(* IEC 61131-3 sources: Industry-PLC-LLM/data/PLCBEAD_repo/PLCBEAD_PLCEmbed-main/PLC-BEAD/Source/PLC_Programs, 701 files *)

(* ---- NETWORK.IEC ---- *)
(*@PROPERTIES_EX@
TYPE: DATA_TYPE
LOCALE: 0
*)
(*----------------------------------------------------------------------------------*)
TYPE

  oscat_NW_BUF_SHORT : ARRAY [0..1407] OF BYTE;
  oscat_NW_BUF_LONG  : ARRAY [0..4095] OF BYTE;

  oscat_NETWORK_BUFFER_SHORT :
  STRUCT
    SIZE   : UINT;
    BUFFER : oscat_NW_BUF_SHORT;
  END_STRUCT;

  oscat_NETWORK_BUFFER :
  STRUCT
    SIZE   : UINT;
    BUFFER : oscat_NW_BUF_LONG;
  END_STRUCT;

END_TYPE

TYPE oscat_url :
    STRUCT
    PROTOCOL : oscat_STRING10;
    USER     : oscat_STRING32;
    PASSWORD : oscat_STRING32;
    DOMAIN   : oscat_STRING80;
    PORT     : WORD;
    PATH     : oscat_STRING80;
    QUERY    : oscat_STRING250;
    ANCHOR   : oscat_STRING40;
    HEADER   : oscat_STRING160;
    END_STRUCT;
END_TYPE

TYPE
  oscat_aB0_5	: ARRAY [0..5] 	OF BYTE;
  oscat_aB0_15	: ARRAY [0..15]	OF BYTE;
  oscat_aB0_19	: ARRAY [0..19]	OF BYTE;
  oscat_aB0_31	: ARRAY [0..31]	OF BYTE;
  oscat_aB0_39	: ARRAY [0..39]	OF BYTE;
  oscat_aB0_47	: ARRAY [0..47]	OF BYTE;
  oscat_aB0_63	: ARRAY [0..63]	OF BYTE;
  oscat_aB0_255	: ARRAY [0..255] OF BYTE;
  oscat_aB1_255	: ARRAY [1..255] OF BYTE;

  oscat_aW0_255	: ARRAY [0..255] OF WORD;
  oscat_aDW0_3	: ARRAY [0..3] 	OF DWORD;
  oscat_aDW0_15	: ARRAY [0..15] OF DWORD;
  oscat_aDW0_4	: ARRAY [0..4] 	OF DWORD;
  oscat_sDW0_79	: ARRAY [0..79] OF DWORD;
END_TYPE

TYPE
  oscat_VMAP_DATA :
  STRUCT
	FC       : DWORD;
    V_ADR    : INT;
    V_SIZE   : INT;
    P_ADR    : INT;
	TIME_OUT : TIME;
  END_STRUCT;

  oscat_MB_VMAP : ARRAY [1..10] OF oscat_VMAP_DATA;

  csv_parser_demo_col : ARRAY [1..4] OF REAL;
  csv_parser_demo     : ARRAY [1..2] OF csv_parser_demo_col;

END_TYPE

TYPE
  oscat_IP_FIFO128_DATA  : ARRAY [1..128] OF BYTE;
  oscat_Mailbox  : ARRAY [1..16] OF BYTE;

  oscat_IP_FIFO_DATA :
  STRUCT
	X       : oscat_IP_FIFO128_DATA; (* IP_ID FIFO Speicher          *)
	Y       : oscat_IP_FIFO128_DATA; (* IP_ID Z�hler                 *)
	ID      : BYTE;                  (* h�chste vergabene id         *)
	MAX_ID  : BYTE;                  (* maximal Anmeldungen pro ID   *)
    INIT    : BOOL;                  (* Initialisierung durchgef�hrt *)
	EMPTY   : BOOL;                  (* FIFO leer                    *)
	FULL    : BOOL;                  (* FIFO voll                    *)
	TOP     : INT;                   (* maximale anzahl in FIFO      *)
	NW      : INT;                   (* Schreibzeiger                *)
	NR      : INT;                   (* Lesezeiger                   *)
  END_STRUCT;

  oscat_IP_C:
  STRUCT
  	C_MODE:			BYTE;          		(*W Mode: TCP/UCP AKTIV/PASSIV                               *)
	C_PORT:         WORD;          		(*W Portnummer                                               *)
	C_IP:           DWORD;         		(*W IP-Adresse gepackt wwxxyyzz = www.xxx.yyy.zzz            *)
    C_STATE:        BYTE;          		(*R Verbindungsstatus ON/OFF + Flanke ON/OFF                 *)
	C_ENABLE:       BOOL;          		(*W Freigabe f�r Connect                                     *)
    R_OBSERVE:      BOOL;          		(*W Empfang ueberwachen                                      *)
    TIME_RESET:     BOOL;          		(*W Alle Timer ruecksetzen                                   *)
	ERROR:          DWORD;         		(*R vvwwxxyy (vv = CON_ERROR, ww = SEN_ERROR, xx = REC_ERROR *)
    FIFO:           oscat_IP_FIFO_DATA; (*I IP FIFO Struktur                                         *)
	MAILBOX:		oscat_Mailbox;		(*I Mailbox: Datenbereich f�r Bausteindatenaustausch         *)
  END_STRUCT;

  oscat_XML_CONTROL:
  STRUCT
    COMMAND:             WORD;            (*W                 *)
    WATCHDOG:            TIME;            (*W                 *)
    START_POS:           UINT;            (*W                 *)
    STOP_POS:            UINT;            (*W                 *)
    COUNT:               UINT;            (*R                 *)
    TYP:                 INT;             (*R                 *)
    LEVEL:               UINT;            (*R                 *)
    PATH:                oscat_STRING250; (*R                 *)
    ELEMENT:             oscat_STRING250; (*R                 *)
    ATTRIBUTE:           oscat_STRING250; (*R                 *)
    VALUE:               oscat_STRING250; (*R                 *)
    BLOCK1_START:        UINT;            (*R                 *)
    BLOCK1_STOP:         UINT;            (*R                 *)
    BLOCK2_START:        UINT;            (*R                 *)
    BLOCK2_STOP:         UINT;            (*R                 *)
  END_STRUCT;

  (* --------- WORLD WEATHER --------- *)

  oscat_WORLD_WEATHER_CUR :
  STRUCT
	OBSERVATION_TIME : oscat_STRING8;
	TEMP_C           : INT;
	WEATHER_CODE     : INT;
	WEATHER_DESC 	 : oscat_STRING60;
	WEATHER_ICON     : INT;
	WIND_SPEED_MILES : INT;
	WIND_SPEED_KMPH  : INT;
	WIND_DIR_DEGREE  : INT;
	WIND_DIR16POINT  : oscat_STRING3;
	PRECIPMM         : REAL;
	HUMIDITY         : INT;
	VISIBILITY       : INT;
	PRESSURE         : INT;
	CLOUDOVER        : INT;
  END_STRUCT;

  oscat_WORLD_WEATHER_DAY :
  STRUCT
	DATE_OF_DAY      : oscat_STRING10;
	TEMP_MAX_C       : INT;
	TEMP_MAX_F       : INT;
	TEMP_MIN_C       : INT;
	TEMP_MIN_F       : INT;
	WIND_SPEED_MILES : INT;
	WIND_SPEED_KMPH  : INT;
	WIND_DIR_DEGREE  : INT;
	WIND_DIR16POINT  : oscat_STRING3;
	WEATHER_CODE     : INT;
	WEATHER_DESC     : oscat_STRING60;
	WEATHER_ICON     : INT;
	PRECIPMM         : REAL;
  END_STRUCT;

  oscat_WORLD_WEATHER_DAY_ARR : ARRAY [0..4] OF oscat_WORLD_WEATHER_DAY;

  oscat_WORLD_WEATHER_DATA :
  STRUCT
	CUR : oscat_WORLD_WEATHER_CUR;
	DAY : oscat_WORLD_WEATHER_DAY_ARR;
  END_STRUCT;

  oscat_WORLD_WEATHER_aI0_41 : ARRAY[0..41] OF INT;

  (* --------- WEATHER CHANNEL --------- *)
  oscat_YAHOO_WEATHER_DATA:
  STRUCT
    TIMETOLIVE:                 INT;              (* TIME TO LIVE: HOW LONG IN MINUTES THIS FEED SHOULD BE CACHED         *)
    LOCATION_CITY:              OSCAT_STRING40;   (* THE LOCATION OF THIS FORECAST: CITY: CITY NAME  *)
    LOCATION_REGION:            OSCAT_STRING20;   (* THE LOCATION OF THIS FORECAST: REGION: STATE, TERRITORY, OR REGION, IF GIVEN *)
    LOCATION_COUNTRY:           OSCAT_STRING20;    (* THE LOCATION OF THIS FORECAST: COUNTRY: TWO-CHARACTER COUNTRY CODE *)
    UNIT_TEMPERATURE:           OSCAT_STRING1;    (* TEMPERATURE: DEGREE UNITS, F FOR FAHRENHEIT OR C FOR CELSIUS *)
    UNIT_DISTANCE:              OSCAT_STRING2;    (* DISTANCE: UNITS FOR DISTANCE, MI FOR MILES OR KM FOR KILOMETERS *)
    UNIT_PRESSURE:              OSCAT_STRING2;    (* PRESSURE: UNITS OF BAROMETRIC PRESSURE, IN FOR POUNDS PER SQUARE INCH OR MB FOR MILLIBARS *)
    UNIT_SPEED:                 OSCAT_STRING4;    (* SPEED: UNITS OF SPEED, MPH FOR MILES PER HOUR OR KPH FOR KILOMETERS PER HOUR *)
    WIND_CHILL:                 INT;              (* FORECAST INFORMATION ABOUT WIND CHILL IN DEGREES *)
    WIND_DIRECTION:             INT;              (* FORECAST INFORMATION ABOUT WIND DIRECTION, IN DEGREES *)
    WIND_SPEED:                 REAL;             (* FORECAST INFORMATION ABOUT WIND SPEED, IN THE UNITS (MPH OR KPH)*)
    ATMOSPHERE_HUMIDITY:        INT;              (* FORECAST INFORMATION ABOUT CURRENT ATMOSPHERIC HUMIDITY: HUMIDITY, IN PERCENT  *)
    ATMOSPHERE_PRESSURE:        INT;              (* FORECAST INFORMATION ABOUT CURRENT ATMOSPHERIC PRESSURE: BAROMETRIC PRESSURE, IN THE UNITS (IN OR MB) *)
	ATMOSPHERE_VISIBILITY:      REAL;             (* FORECAST INFORMATION ABOUT CURRENT ATMOSPHERIC VISIBILITY, IN THE UNITS (MI OR KM) *)
	ATMOSPHERE_RISING:          INT;              (* FORECAST INFORMATION ABOUT RISING: STATE OF THE BAROMETRIC PRESSURE: STEADY (0), RISING (1), OR FALLING (2). (INTEGER: 0, 1, 2) *)
    ASTRONOMY_SUNRISE:          OSCAT_STRING10;   (* SUNRISE: TODAY'S SUNRISE TIME. THE TIME IS A STRING IN A LOCAL TIME FORMAT OF "H:MM AM/PM" *)
    ASTRONOMY_SUNSET:           OSCAT_STRING10;   (* SUNSET: TODAY'S SUNSET TIME. THE TIME IS A STRING IN A LOCAL TIME FORMAT OF "H:MM AM/PM", *)
    GEO_LATITUDE:               REAL;             (* THE LATITUDE OF THE LOCATION *)
    GEO_LONGITUDE:              REAL;             (* THE LONGITUDE OF THE LOCATION *)
    CUR_CONDITIONS_TEMP:        INT;              (* THE CURRENT WEATHER CONDITIONS: TEMP: THE CURRENT TEMPERATURE, IN THE UNITS (F OR C) *)
    CUR_CONDITIONS_TEXT:        OSCAT_STRING40;   (* THE CURRENT WEATHER CONDITIONS: TEXT: A TEXTUAL DESCRIPTION OF CONDITIONS *)
    CUR_CONDITIONS_CODE:        INT;              (* THE CURRENT WEATHER CONDITIONS: CODE: THE CONDITION CODE FOR THIS FORECAST *)
	CUR_CONDITIONS_ICON:        INT;			  (* THE CURRENT WEATHER CONDITIONS: ICON: THE CONDITION ICON FOR THIS FORECAST *)
    FORCAST_TODAY_LOW_TEMP:     INT;              (* THE FORCAST TODAY WEATHER CONDITIONS: THE FORECASTED LOW TEMPERATURE FOR THIS DAY IN THE UNITS (F OR C) *)
    FORCAST_TODAY_HIGH_TEMP:    INT;              (* THE FORCAST TODAY WEATHER CONDITIONS: THE FORECASTED HIGH TEMPERATURE FOR THIS DAY IN THE UNITS (F OR C) *)
    FORCAST_TODAY_TEXT:         OSCAT_STRING40;   (* THE FORCAST TODAY WEATHER CONDITIONS: TEXT: A TEXTUAL DESCRIPTION OF CONDITIONS *)
    FORCAST_TODAY_CODE:         INT;              (* THE CURRENT WEATHER CONDITIONS: CODE: THE CONDITION CODE FOR THIS FORECAST *)
	FORCAST_TODAY_ICON:         INT;			  (* THE CURRENT WEATHER CONDITIONS: ICON: THE CONDITION ICON FOR THIS FORECAST *)
    FORCAST_TOMORROW_LOW_TEMP:  INT;              (* THE FORCAST TOMORROW WEATHER CONDITIONS: THE FORECASTED LOW TEMPERATURE FOR THIS DAY IN THE UNITS (F OR C) *)
    FORCAST_TOMORROW_HIGH_TEMP: INT;              (* THE FORCAST TOMORROW WEATHER CONDITIONS: THE FORECASTED HIGH TEMPERATURE FOR THIS DAY IN THE UNITS (F OR C) *)
    FORCAST_TOMORROW_TEXT:      OSCAT_STRING40;   (* THE FORCAST TOMORROW WEATHER CONDITIONS: TEXT: A TEXTUAL DESCRIPTION OF CONDITIONS *)
    FORCAST_TOMORROW_CODE:      INT;              (* THE CURRENT WEATHER CONDITIONS: CODE: THE CONDITION CODE FOR THIS FORECAST *)
	FORCAST_TOMORROW_ICON:      INT;			  (* THE CURRENT WEATHER CONDITIONS: ICON: THE CONDITION ICON FOR THIS FORECAST *)
  END_STRUCT;

  oscat_YAHOO_WEATHER_aI0_48 : ARRAY[0..48] OF INT;

  oscat_IP2GEO_DATA:
  STRUCT
	STATE :				BOOL;			  (* STATE *)
	IP4 :				DWORD;			  (* IP-Adresse *)
    COUNTRY_CODE :		oscat_STRING2;    (*   *)
    COUNTRY_NAME :		oscat_STRING20;   (*   *)
    REGION_CODE :		oscat_STRING2;    (*   *)
    REGION_NAME :		oscat_STRING20;   (*   *)
    CITY :				oscat_STRING20;   (*   *)
    GEO_LATITUDE :		REAL;             (*   *)
    GEO_LONGITUDE :		REAL;             (*   *)
	TIME_ZONE_NAME :	oscat_STRING20;
	GMT_OFFSET :		INT;
	IS_DST :			BOOL;
  END_STRUCT;
END_TYPE

(*----------------------------------------------------------------------------------*)

TYPE
  PRINTF_DATA_250  	:  ARRAY [1..11]  OF oscat_STRING250;
  PRINTF_DATA_80 	:  ARRAY [1..11]  OF oscat_STRING80;
  LOG_250       	:  ARRAY [0..400] OF oscat_STRING250;
  LOG_80    		:  ARRAY [0..400] OF oscat_STRING80;
  LOG_OPTION		:  ARRAY [0..400] OF DWORD;

  us_LOG_CONTROL :
  STRUCT
    NEW_MSG              : oscat_STRING250;    (*W neue Nachricht f�r den Datenbuffer   *)
	NEW_MSG_OPTION 		 : DWORD;
    LEVEL                : BYTE;
	SIZE                 : INT;                (*R Anzahl der Strings im LOG_DATA       *)
	RESET                : BOOL;               (*W Nachrichtenbuffer l�schen            *)
    PRINTF               : PRINTF_DATA_250;    (*W Array PRINTF Parameter               *)
    MSG                  : LOG_250;            (*I Array Message                        *)
    MSG_OPTION           : LOG_OPTION;     	   (*I Array Message Option                 *)
	UPDATE_COUNT         : UINT;               (*R Updatez�hler                         *)
    IDX                  : INT;                (*R aktueller Nachrichten-Index          *)
	RING_MODE            : BOOL;               (*I Buffer�berlauf erkannt               *)
  END_STRUCT;

  us_LOG_CONTROL_80 :
  STRUCT
    NEW_MSG              : oscat_STRING80;     (*W neue Nachricht f�r den Datenbuffer   *)
	NEW_MSG_OPTION 		 : DWORD;
    LEVEL                : BYTE;
	SIZE                 : INT;                (*R Anzahl der Strings im LOG_DATA       *)
	RESET                : BOOL;               (*W Nachrichtenbuffer l�schen            *)
    PRINTF               : PRINTF_DATA_80;     (*W Array PRINTF Parameter               *)
    MSG                  : LOG_80;             (*I Array Message                        *)
    MSG_OPTION           : LOG_OPTION;     	   (*I Array Message Option                 *)
	UPDATE_COUNT         : UINT;               (*R Updatez�hler                         *)
    IDX                  : INT;                (*R aktueller Nachrichten-Index          *)
	RING_MODE            : BOOL;               (*I Buffer�berlauf erkannt               *)
  END_STRUCT;

  LINE_ARRAY 			: ARRAY [1..40] OF INT;

  us_LOG_VIEWPORT :
    STRUCT
     LINE_ARRAY          : LINE_ARRAY;
     COUNT               : INT;                (* Anzahl der sichtbaren Nachtrichten   *)
	 UPDATE_COUNT        : UINT;               (* Updatez�hler                         *)
     MOVE_TO_X           : INT;                (* Steuerung der Nachrichtenanzeige     *)
     UPDATE              : BOOL;               (* Daten wurden ge�ndert -> neuzeichnen *)
  END_STRUCT;

  oscat_FILE_SERVER_DATA : STRUCT
	FILE_OPEN	: BOOL;
    FILENAME 	: STRING;
    MODE	 	: BYTE;
    OFFSET   	: UDINT;
    FILE_SIZE   : UDINT;
    AUTO_CLOSE	: TIME;
    ERROR	 	: BYTE;
  END_STRUCT;

  oscat_FILE_PATH_DATA : STRUCT
	DRIVE : oscat_string3;
	DIRECTORY : oscat_string250;
	FILENAME : STRING;
  END_STRUCT;

  oscat_UNI_CIRCULAR_BUFFER_DATA : STRUCT
	D_MODE : INT;
	D_HEAD : WORD;
	D_STRING : oscat_string250;
	D_REAL : REAL;
	D_DWORD : DWORD;
	BUF_SIZE : INT;
	BUF_COUNT : INT;
	BUF_USED : USINT;
	BUF : oscat_NW_BUF_LONG;
	_GetStart : INT;
	_GetEnd : INT;
	_Last : INT;
	_First : INT;
  END_STRUCT;

  oscat_DLOG_DATA : STRUCT
	STORE_TYPE : BYTE;
	ADD_HEADER : BOOL;
	ADD_DATA : BOOL;
	ADD_DATA_REQ : BOOL;
	CLOCK_TRIG : BOOL;
	ID_MAX : USINT;
	DTI : UDINT;
	UCB : oscat_UNI_CIRCULAR_BUFFER_DATA;
	NEW_FILE : STRING;
	NEW_FILE_RTRIG : BOOL;
  END_STRUCT;

END_TYPE
(* --------------------------- NET_VAR ---------------------------- *)
TYPE oscat_NET_VAR_DATA :
STRUCT
	CYCLE : UDINT;
	STATE : BYTE;
	INDEX : INT;
	ID_MAX : USINT;
	ERROR_ID : BYTE;
	BUF_SIZE : UINT;
	S_BUF : oscat_NETWORK_BUFFER;
	R_BUF : oscat_NETWORK_BUFFER;
END_STRUCT;
END_TYPE

TYPE
    oscat_aB1_64 : ARRAY[1..64] OF BYTE;
	oscat_nv_ra : ARRAY[1..8] OF REAL;
	oscat_nv_dw : ARRAY[1..8] OF DWORD;
END_TYPE

(* --------------------------- TELNET ----------------------------- *)

TYPE

(*----------------------------------------------------------------------------------*)
(* Menue-System                                                                     *)
(*----------------------------------------------------------------------------------*)

  us_TN_MENU_POPUP :
  STRUCT
    st_Menu_Text:         oscat_STRING250;   (* X Menue Texte                               *)
    in_Menu_E_Count:      INT;               (*   Menue Elemente Anzahl                     *)
    in_X:                 INT;               (* X Menue X-Position                          *)
    in_Y:                 INT;               (* X Menue Y-Position                          *)
    in_Cols:              INT;               (*   Menue Spaltenanzahl                       *)
    in_Rows:              INT;               (*   Menue Zeilenanzahl                        *)
    in_Cur_Item:          INT;               (* X aktuelles Sub-Menue                       *)
    by_Attr_mF:           BYTE;              (* X Text Attribute mit Fokus                  *)
    by_Attr_oF:           BYTE;              (* X Text Attribute ohne Fokus                 *)
    by_Input_Exten_Code:  BYTE;              (* X Tastencode: Sondertasten                  *)
    bo_Create:            BOOL;              (* X Popup-Menu erzeugen                       *)
    bo_Destroy:           BOOL;              (* X Popup-Menu entfernen                      *)
    bo_Update:            BOOL;              (* X Popup-Menu updaten                        *)
    bo_Activ:             BOOL;              (*   Popup-Menu ist aktiv                      *)
  END_STRUCT;

  us_TN_MENU :
  STRUCT
    st_Menu_Text:         oscat_STRING250;   (* X Menue Texte                               *)
    in_Menu_E_Count:      INT;               (* Menue Elemente Anzahl                       *)
    in_Y:                 INT;               (* Menue Zeilennummer  Y-Position              *)
    in_X:                 INT;               (* Menue Spaltennummer X-Position              *)
    by_Attr_mF:           BYTE;              (* Text Attribute mit Fokus                    *)
    by_Attr_oF:           BYTE;              (* Text Attribute ohne Fokus                   *)
    in_X_SM_new:          INT;               (* neue Sub-Menu X-Position                    *)
    in_Y_SM_new:          INT;               (* neue Sub-Menu Y-Position                    *)
    in_X_SM_old:          INT;               (* alte Sub-Menu X-Position                    *)
    in_Y_SM_old:          INT;               (* alte Sub-Menu Y-Position                    *)
    in_Cur_Menu_Item:     INT;               (* aktuelles Haupt-Menue                       *)
    in_Cur_Sub_Item:      INT;               (* aktuelles Sub-Menue                         *)
    in_State:             INT;               (*   Menu status                               *)
    in_Menu_Selected:     INT;               (* X Menu-Item mit Enter angew�hlt             *)
    bo_Create:            BOOL;              (* X Menu erzeugen                             *)
    bo_Destroy:           BOOL;              (* X Menu entfernen                            *)
    bo_Update:            BOOL;              (* X Menu updaten                              *)

  END_STRUCT;

(*----------------------------------------------------------------------------------*)

  bya_TN_CHAR:       	ARRAY [0..1919] OF BYTE;
  bya_TN_BACKUP:     	ARRAY [0..1919] OF BYTE;
  bya_TN_COLOR:      	ARRAY [0..1919] OF BYTE;
  bya_TN_Line_Update:	ARRAY [0..23]   OF BOOL;

  us_TN_SCREEN :
  STRUCT
    bya_CHAR:			bya_TN_CHAR;
    bya_COLOR:			bya_TN_COLOR;
    bya_BACKUP:			bya_TN_BACKUP;
    bya_Line_Update:	bya_TN_Line_Update;

    by_Input_Exten_Code:    BYTE;
    by_Input_ASCII_Code:    BYTE;
    bo_Input_ASCII_IsNum:   BOOL;
    in_Page_Number:        	INT;                (* aktive Seiten-Nr.              *)
    in_Cursor_X:           	INT;                (* Cursor X-Position              *)
    in_Cursor_Y:           	INT;                (* Cursor Y-Position              *)
    in_EOS_Offset:         	INT;                (* End of String Offset           *)
    by_Clear_Screen_Attr:  	BYTE;               (* Clear-Screen Attr              *)
    bo_Clear_Screen:       	BOOL;               (* Clear-Screen ausl�sen          *)
    bo_Modal_Dialog:       	BOOL;               (* Modaler Dialog ist aktiv       *)
    bo_Menue_Bar_Dialog:   	BOOL;               (* Menue Dialog ist aktiv         *)

  END_STRUCT;

(*----------------------------------------------------------------------------------*)

  us_TN_INPUT_CONTROL_DATA :
  STRUCT
    by_Input_Exten_Code:    BYTE;
    by_Input_ASCII_Code:    BYTE;
    bo_Input_ASCII_IsNum:   BOOL;
    in_Title_X_Offset:  	INT;         	(* Title Text X-Offset                       *)
    in_Title_Y_Offset:   	INT;         	(* Title Text Y-Offset                       *)
    by_Title_Attr:			BYTE;        	(* Title Text Attribute                      *)
    st_Title_String:    	STRING;      	(* Title Text String                         *)
    in_Cursor_X:          	INT;			(* aktuelle Cursor X-Position                *)
    in_Cursor_Y:          	INT;			(* aktuelle Cursor Y-Position                *)
    in_Type:              	INT;            (* Type des Elements                         *)
    in_X:                 	INT;            (* Element X-Position                        *)
    in_Y:                 	INT;            (* Element Y-Position                        *)
    in_Cursor_Pos:        	INT;            (* aktuelle Cursorposition                   *)
    by_Attr_mF:           	BYTE;           (* Text Attribute mit Fokus                  *)
    by_Attr_oF:           	BYTE;           (* Text Attribute ohne Fokus                 *)
	in_selected:          	INT;            (* Text Item wurde ausgew�hlt                *)
    st_Input_Mask:        	STRING;         (* Text Eingabemaske                         *)
    st_Input_Data:        	oscat_STRING250;(* Text aktuelle Eingabedaten                *)
    st_Input_String:      	STRING;         (* Text Kopie nach Return-Taste              *)
    st_Input_ToolTip:     	STRING;         (* Text ToolTip (Eingabeinformation)         *)
	in_Input_Option:      	INT;            (* Text Ausgabe-Optionen                     *)
	bo_Input_Entered:     	BOOL;           (* RETURN-Taste wurde bet�tigt               *)
    bo_Input_Hidden:      	BOOL;           (* Text versteckete Eingabe mit '*'          *)
	bo_Input_Only_Num:    	BOOL;           (* Text nur Nummerneingabe zulassen          *)
	bo_Focus:             	BOOL;           (* Element besitzt den Fokus                 *)
	bo_Update_Input:      	BOOL;           (* Element wegen Benutzereingabe neuzeichnen *)
	bo_Update_All:        	BOOL;           (* Element komplett neuzeichnen              *)

  END_STRUCT;

  usa_TN_INPUT_CONTROL_DATA:   ARRAY [1..20] OF us_TN_INPUT_CONTROL_DATA;

  us_TN_INPUT_CONTROL :
  STRUCT
    bo_Enable:          BOOL;           (* Bearbeitung freigeben/sperren           *)
    bo_Update_all:      BOOL;           (* All Elemente neu zeichnen               *)
    bo_Reset_Fokus:     BOOL;           (* Fokus auf 1. Element setzen             *)
    in_Focus_at:        INT;            (* Controlelement mit aktivem Fokus        *)
    in_Count:           INT;            (* Anzahl der benutzen Control-Elemente    *)
    in_ToolTip_X:       INT;            (* Tooltip Text X-Offset                   *)
    in_ToolTip_Y:		INT;            (* Tooltip Text Y-Offset                   *)
    by_ToolTip_Attr:	BYTE;           (* Tooltip Text Attribute                  *)
    in_ToolTip_Size:	INT;            (* Tooltip Text l�nge                      *)
    usa_TN_INPUT_CONTROL_DATA: usa_TN_INPUT_CONTROL_DATA;
  END_STRUCT;

END_TYPE

(* ---- OSCAT.IEC ---- *)
(*@PROPERTIES_EX@
TYPE: DATA_TYPE
LOCALE: 0
*)
TYPE
  oscat_STRING1               : STRING(1);
  oscat_STRING2               : STRING(2);
  oscat_STRING3               : STRING(3);
  oscat_STRING4               : STRING(4);
  oscat_STRING5               : STRING(5);
  oscat_STRING8               : STRING(8);
  oscat_STRING10              : STRING(10);
  oscat_STRING12              : STRING(12);
  oscat_STRING15              : STRING(15);
  oscat_STRING20              : STRING(20);
  oscat_STRING27              : STRING(27);
  oscat_STRING30              : STRING(30);
  oscat_STRING32              : STRING(32);
  oscat_STRING40              : STRING(40);
  oscat_STRING48              : STRING(48);
  oscat_STRING50              : STRING(50);
  oscat_STRING60              : STRING(60);
  oscat_STRING64              : STRING(64);
  oscat_STRING80              : STRING(80);
  oscat_STRING120             : STRING(120);
  oscat_STRING144             : STRING(144);
  oscat_STRING160             : STRING(160);
  oscat_STRING189             : STRING(189);
  oscat_STRING192             : STRING(192);
  oscat_STRING250             : STRING(250);
END_TYPE

(*----------------------------------------------------------------------------------*)
TYPE

  oscat_arr_0_7               : ARRAY [0..7]    OF REAL;
  oscat_arr_0_15              : ARRAY [0..15]   OF REAL;
  oscat_delay_buf             : ARRAY [0..31]   OF REAL;
  oscat_FT_TN64_array         : ARRAY [0..63]   OF REAL;
  oscat_pt_ARRAY              : ARRAY [1..100]  OF REAL;

  oscat_ardw_0_15             : ARRAY [0..15]   OF DWORD;
  oscat_ardw_0_31             : ARRAY [0..31]   OF DWORD;

  oscat_FILTER_MAV_W          : ARRAY [0..31]   OF WORD;
  oscat_arb_0_3               : ARRAY [0..3]    OF BYTE;

  oscat_esr_collect_data      : ARRAY [0..7]    OF BYTE;
  oscat_DRIVER_4C 			  : ARRAY [1..7] 	OF BYTE;
  oscat_arb_0_249 			  : ARRAY [0..249] 	OF BYTE;
  oscat_bya_LIST_CLEAN        : ARRAY [1..250]  OF BYTE;

  oscat_ari_0_30         	  : ARRAY [0..30]   OF INT;

  oscat_stack_array 		  : ARRAY [1..32]   OF INT;

  oscat_dcf77_bits            : ARRAY [0..58]   OF BOOL;

  oscat_array64_time          : ARRAY [0..63]   OF TIME;

  (* -------------------------------------------------- *)
  oscat_PERIOD2_Y             : ARRAY [0..1]    OF UDINT;
  oscat_PERIOD2_X             : ARRAY [0..3]    OF oscat_PERIOD2_Y;

  oscat_ARRAY_X               : ARRAY [0..1]    OF REAL;
  oscat_XY                    : ARRAY [1..20]   OF oscat_ARRAY_X;

  oscat_parset_X              : ARRAY [1..4]    OF REAL;
  oscat_parset                : ARRAY [0..3]    OF oscat_parset_X;

  oscat_Polynom_ARRAY_X       : ARRAY [0..1]    OF REAL;
  oscat_Polynom_XY            : ARRAY [1..5]    OF oscat_Polynom_ARRAY_X;

END_TYPE

(*----------------------------------------------------------------------------------*)
TYPE oscat_FRACTION :
STRUCT
	NUMERATOR : INT;
	DENOMINATOR : INT;
END_STRUCT;
END_TYPE
(*----------------------------------------------------------------------------------*)
TYPE oscat_CALENDAR :
	STRUCT
		UTC : UDINT;				(* world time UTC *)
		LDT : UDINT;				(* local time *)
		LDATE : UDINT;				(* local date *)
		LTOD : UDINT;				(* local time of day *)
		YEAR : INT;					(* year of LDATE *)
		MONTH : INT;				(* month of LDATE *)
		DAY : INT;					(* day of LDATE *)
		WEEKDAY : INT;				(* weekday of LDATE *)
		OFFSET : INT;				(* Time Zone Offset for Local time in minutes *)
		DST_EN : BOOL;				(* daylight savings time enable *)
		DST_ON : BOOL;				(* true when daylight savings time os on *)
		NAME : oscat_string5;		(* name of time zone *)
		LANGUAGE : INT;			    (* language number pls see language setup *)
		LONGITUDE : REAL;			(* longitude of current location *)
		LATITUDE : REAL;			(* latitude of current location *)
		SUN_RISE : UDINT;			(* sun_rise for current location *)
		SUN_SET : UDINT;			(* sun_set for current location *)
		SUN_MIDDAY : UDINT;			(* worldtime when sun stands at south position *)
		SUN_HEIGTH : REAL;			(* suns heigth at midday, south position *)
		SUN_HOR : REAL;				(* sun angle horizontal 0 = north in degrees *)
		SUN_VER : REAL;				(* sun angle vertical above horizon in degrees *)
		NIGHT : BOOL;				(* true between sun_set and sun_rise *)
		HOLIDAY : BOOL;				(* true when holiday *)
		HOLY_NAME : oscat_string30;	(* name of holiday *)
		WORK_WEEK : INT;			(* current work week *)
	END_STRUCT;
END_TYPE

TYPE oscat_SDT :
STRUCT
	YEAR : INT;
	MONTH : INT;
	DAY : INT;
	WEEKDAY : INT;
	HOUR : INT;
	MINUTE : INT;
	SECOND : INT;
	MS : INT;
END_STRUCT;
END_TYPE

(*----------------------------------------------------------------------------------*)

TYPE oscat_LANGUAGE:
  STRUCT
    DEFAULT 	: INT;
	LMAX    	: INT;
  END_STRUCT;
END_TYPE

(*----------------------------------------------------------------------------------*)
TYPE
	oscat_LOCATION_ELEMENTS	: ARRAY [1..5] OF INT;
END_TYPE

TYPE oscat_LOCATION:
  STRUCT
    DEFAULT 	: INT;
	LMAX    	: INT;
	LANGUAGE	: oscat_LOCATION_ELEMENTS;
  END_STRUCT;
END_TYPE

(*----------------------------------------------------------------------------------*)

TYPE
  oscat_ELEMENT_DIRS 		: ARRAY [0..15] OF oscat_STRING3;
  oscat_DIRS				: ARRAY [1..3]  OF oscat_ELEMENT_DIRS;
END_TYPE

(*----------------------------------------------------------------------------------*)
TYPE
  oscat_CHARNAMES	: ARRAY [1..11] OF STRING;
END_TYPE

(*----------------------------------------------------------------------------------*)

TYPE
  oscat_ELEMENT_MONTHS 	: ARRAY [1..12] OF oscat_STRING10;
  oscat_MONTHS			: ARRAY [1..3]  OF oscat_ELEMENT_MONTHS;
END_TYPE

(*----------------------------------------------------------------------------------*)

TYPE
  oscat_ELEMENT_MONTHS3	: ARRAY [1..12] OF oscat_STRING3;
  oscat_MONTHS3			: ARRAY [1..3]  OF oscat_ELEMENT_MONTHS3;
END_TYPE

(*----------------------------------------------------------------------------------*)

TYPE
  oscat_ELEMENT_WEEKDAYS	: ARRAY [1..7] OF oscat_STRING10;
  oscat_WEEKDAYS			: ARRAY [1..3]  OF oscat_ELEMENT_WEEKDAYS;
END_TYPE

(*----------------------------------------------------------------------------------*)

TYPE
  oscat_ELEMENT_WEEKDAYS2	: ARRAY [1..7] OF oscat_STRING2;
  oscat_WEEKDAYS2			: ARRAY [1..3]  OF oscat_ELEMENT_WEEKDAYS2;
END_TYPE

TYPE oscat_esr_data :
  STRUCT
	typ    : BYTE;
	adress : oscat_string10;
	DS     : UDINT;
	TS     : TIME;
	data   : oscat_esr_collect_data;
  END_STRUCT;
END_TYPE

TYPE
  oscat_ESR_3                : ARRAY [0..3] OF oscat_esr_data;
  oscat_ESR_31               : ARRAY [0..31] OF oscat_esr_data;
END_TYPE

TYPE oscat_vector_3 :
  STRUCT
	X : REAL;
	Y : REAL;
	Z : REAL;
  END_STRUCT;
END_TYPE

TYPE oscat_complex :
  STRUCT
	re : REAL;
	im : REAL;
  END_STRUCT;
END_TYPE

TYPE REAL2 :
  STRUCT
	R1 : REAL;
	RX : REAL;
  END_STRUCT;
END_TYPE

(*----------------------------------------------------------------------------------*)

TYPE oscat_HOLIDAY_DATA :
  STRUCT
	NAME : oscat_string30;
	DAY : SINT;
	MONTH : SINT;
	USE : SINT;
	PAD_BYTE : BYTE;
  END_STRUCT;
END_TYPE

TYPE
  oscat_HOLIDAY_DATA_0_29 	: ARRAY [0..29] OF oscat_HOLIDAY_DATA;
  oscat_HOLIDAY_DATA_0_49 	: ARRAY [0..49] OF oscat_HOLIDAY_DATA;
END_TYPE

(* revision history
hm	18. oct. 2008
	original version

*)

(*	if month = 0 then F_day is the offset in days from easter
	used :0 = NOT used, 1 = used, -1..-7 menas the weekday before the specified DATE example -3 means wednesday before 23.11
*)

(* samples for Holiday data

	HOLIDAY_DE : ARRAY[0..29] OF HOLIDAY_DATA := (name := 'Neujahr', day := 1, month := 1, use := 1),
		(name := 'Heilig Drei Könige', day := 6, month := 1, use := 1),
		(name := 'Karfreitag', day := -2, month := 0, use := 1),
		(name := 'Ostersonntag', day := 0, month := 0, use := 1),
		(name := 'Ostermontag', day := 1, month := 0, use := 1),
		(name := 'Tag der Arbeit', day := 1, month := 5, use := 1),
		(name := 'Christi Himmelfahrt', day := 39, month := 0, use := 1),
		(name := 'Pfingstsonntag', day := 49, month := 0, use := 1),
		(name := 'Pfingstmontag', day := 50, month := 0, use := 1),
		(name := 'Fronleichnam', day := 60, month := 0, use := 1),
		(name := 'Augsburger Friedensfest', day := 8, month := 8, use := 0),
		(name := 'Maria Himmelfahrt', day := 15, month := 8, use := 1),
		(name := 'Tag der Deutschen Einheit', day := 3, month := 10, use := 1),
		(name := 'Reformationstag', day := 31, month := 10, use := 0),
		(name := 'Allerheiligen', day := 1, month := 11, use := 1),
		(name := 'Buss und Bettag', day := 23, month := 11, use := 0),
		(name := '1. Weihnachtstag', day := 25, month := 12, use := 1),
		(name := '2. Weihnachtstag', day := 26, month := 12, use := 1);

	HOLIDAY_AT : ARRAY[0..29] OF HOLIDAY_DATA := (name := 'Neujahr', day := 1, month := 1, use := 1),
		(name := 'Heilig Drei Könige', day := 6, month := 1, use := 1),
		(name := 'Karfreitag', day := -2, month := 0, use := 1),
		(name := 'Ostersonntag', day := 0, month := 0, use := 1),
		(name := 'Ostermontag', day := 1, month := 0, use := 1),
		(name := '', day := 1, month := 5, use := 0),
		(name := 'Christi Himmelfahrt', day := 39, month := 0, use := 1),
		(name := 'Pfingstsonntag', day := 49, month := 0, use := 1),
		(name := 'Pfingstmontag', day := 50, month := 0, use := 1),
		(name := 'Fronleichnam', day := 60, month := 0, use := 1),
		(name := '', day := 8, month := 8, use := 0),
		(name := 'Maria Himmelfahrt', day := 15, month := 8, use := 1),
		(name := '', day := 3, month := 10, use := 0),
		(name := '', day := 31, month := 10, use := 0),
		(name := 'Allerheiligen', day := 1, month := 11, use := 1),
		(name := 'Maria Empfängnis', day := 8, month := 12, use := 1),
		(name := '1. Weihnachtstag', day := 25, month := 12, use := 1),
		(name := '2. Weihnachtstag', day := 26, month := 12, use := 1);

	HOLIDAY_FR : ARRAY[0..29] OF HOLIDAY_DATA := (name := 'Nouvel an', day := 1, month := 1, use := 1),
		(name := 'St Valentin', day := 14, month := 2, use := 0),
		(name := 'Vendredi Saint (alsace)', day := -2, month := 0, use := 0),
		(name := 'Dimanche de pâques', day := 0, month := 0, use := 1),
		(name := 'Lundi de pâques', day := 1, month := 0, use := 1),
		(name := 'Jeudi de Ascension', day := 39, month := 0, use := 1),
		(name := 'dimanche de Pentecôte ', day := 49, month := 0, use := 1),
		(name := 'jeudi de la Trinité', day := 60, month := 0, use := 0),
		(name := 'Fête du travail', day := 1, month := 5, use := 1),
		(name := 'Victoire 1945 ', day := 8, month := 5, use := 1),
		(name := 'Prise de La bastille', day := 14, month := 7, use := 1),
		(name := '15 Août 1944', day := 15, month := 8, use := 1),
		(name := 'Halloween', day := 31, month := 10, use := 0),
		(name := 'Armistice 1918', day := 11, month := 11, use := 1),
		(name := 'Noël', day := 25, month := 12, use := 1),
		(name := 'Saint Étienne (alsace)', day := 26, month := 12, use := 0),
		(name := 'Fête de la musique', day := 21, month := 6, use := 0);

	HOLIDAY_BED : ARRAY[0..29] OF HOLIDAY_DATA :=	(name := 'Neujahr', day := 1, month := 1, use := 1),
		(name := 'Ostersonntag', day := 0, month := 0, use := 1),
		(name := 'Ostermontag', day := 1, month := 0, use := 1),
		(name := 'Tag der Arbeit', day := 1, month := 5, use := 1),
		(name := 'Christi Himmelfahrt', day := 39, month := 0, use := 1),
		(name := 'Pfingsten', day := 49, month := 0, use := 1),
		(name := 'Pfingstmontag', day := 50, month := 0, use := 1),
		(name := 'Nationalfeiertag', day := 21, month := 7, use := 1),
		(name := 'Mariä Himmelfahrt', day := 15, month := 8, use := 1),
		(name := 'Allerheiligen', day := 1, month := 11, use := 1),
		(name := 'Feiertag DG', day := 15, month := 11, use := 1),
		(name := 'Heiligabend', day := 24, month := 12, use := 1),
		(name := '1. Weihnachtstag', day := 25, month := 12, use := 1),
		(name := '2. Weihnachtstag', day := 26, month := 12, use := 1),
		(name := 'Silvester', day := 31, month := 12, use := 1);

	HOLIDAY_ITD : ARRAY[0..29] OF HOLIDAY_DATA := (name := 'Neujahr', day := 1, month := 1, use := 1),
		(name := 'Heilig Drei Könige', day := 6, month := 1, use := 1),
		(name := 'Ostersonntag', day := 0, month := 0, use := 1),
		(name := 'Ostermontag', day := 1, month := 0, use := 1),
		(name := 'Tag der Befeiung Italiens', day := 25, month := 4, use := 1),
		(name := 'Tag der Arbeit', day := 1, month := 5, use := 1),
		(name := 'Pfingsten', day := 49, month := 0, use := 1),
		(name := 'Pfingstmontag', day := 50, month := 0, use := 1),
		(name := 'Tag der Republik Italien', day := 2, month := 6, use := 1),
		(name := 'Mariä Himmelfahrt', day := 15, month := 8, use := 1),
		(name := 'Allerheiligen', day := 1, month := 11, use := 1),
		(name := 'Mariä Empfängnis', day := 8, month := 12, use := 1),
		(name := 'Heiligabend', day := 24, month := 12, use := 0),
		(name := '1. Weihnachtstag', day := 25, month := 12, use := 1),
		(name := '2. Stephanstag', day := 26, month := 12, use := 1);

*)

(* ---- TIMER_P4.ST ---- *)
TYPE oscat_TIMER_EVENT_DATA :
  STRUCT
	TYP          : BYTE;
	CHANNEL      : BYTE;
	DAY          : BYTE;
	START        : UDINT;
	DURATION     : TIME;
	LAND         : BYTE;
	LOR          : BYTE;
	LAST         : UDINT;
  END_STRUCT;
END_TYPE

TYPE
  oscat_TIMER_EVENT           : ARRAY [0..63]    OF oscat_TIMER_EVENT_DATA;
  oscat_TP4_qn                : ARRAY [0..3]    OF BOOL;
END_TYPE

TYPE
  oscat_arb_0_3               : ARRAY [0..3]    OF BYTE;
END_TYPE

FUNCTION _BYTE_TO_INT:INT
	VAR_INPUT
		IN :	BYTE;
	END_VAR

	_BYTE_TO_INT := USINT_TO_INT(BYTE_TO_USINT(IN));
END_FUNCTION

FUNCTION DATE_TO_DT:UDINT
	VAR_INPUT
		IN :	UDINT;
	END_VAR
	DATE_TO_DT := IN;
END_FUNCTION

FUNCTION _DT_TO_DATE_B:UDINT

	VAR_INPUT
		_INN :	UDINT;
	END_VAR

	_DT_TO_DATE_B := (_INN / UDINT#86400) * UDINT#86400;
END_FUNCTION

FUNCTION TIME_TO_UDINT2:UDINT
	VAR_INPUT
		X :	TIME;
	END_VAR

	TIME_TO_UDINT2 := DINT_TO_UDINT(TIME_TO_DINT(X));
END_FUNCTION

FUNCTION DATE_TO_UDINT2:UDINT
	VAR_INPUT
		IN :	UDINT;
	END_VAR

	DATE_TO_UDINT2 := IN;
END_FUNCTION

FUNCTION DAY_OF_WEEK:INT
  VAR_INPUT
    IDATE :	UDINT;
  END_VAR

  DAY_OF_WEEK := UDINT_TO_INT((idate / UDINT#86400 + UDINT#3) MOD UDINT#7) + INT#01;
END_FUNCTION

FUNCTION _BYTE_TO_DINT:DINT
	VAR_INPUT
		IN :	BYTE;
	END_VAR

	_BYTE_TO_DINT := USINT_TO_DINT(BYTE_TO_USINT(IN));
END_FUNCTION

FUNCTION DAY_OF_YEAR_UDINT:INT
	VAR_INPUT
		IDATE :	UDINT;
	END_VAR

	DAY_OF_YEAR_UDINT := UDINT_TO_INT((idate / UDINT#86400) MOD UDINT#1461);
	IF DAY_OF_YEAR_UDINT > 729 THEN
		IF DAY_OF_YEAR_UDINT > 1095 THEN DAY_OF_YEAR_UDINT := DAY_OF_YEAR_UDINT - 1095; ELSE DAY_OF_YEAR_UDINT := DAY_OF_YEAR_UDINT - 729; END_IF;
	ELSIF DAY_OF_YEAR_UDINT > 364 THEN
		DAY_OF_YEAR_UDINT := DAY_OF_YEAR_UDINT - 364;
	ELSE
		DAY_OF_YEAR_UDINT := DAY_OF_YEAR_UDINT + 1;
	END_IF;
END_FUNCTION

FUNCTION MONTH_OF_DATE_UDINT:INT

	VAR_INPUT
		IDATE :	UDINT;
	END_VAR

	MONTH_OF_DATE_UDINT := DAY_OF_YEAR_UDINT(idate);
	IF MONTH_OF_DATE_UDINT < 32 THEN
		MONTH_OF_DATE_UDINT := 1;
	ELSIF LEAP_OF_DATE(IDATE) THEN
		MONTH_OF_DATE_UDINT := (MONTH_OF_DATE_UDINT * 53 + 1668) / 1623;
	ELSE
		MONTH_OF_DATE_UDINT := (MONTH_OF_DATE_UDINT * 53 + 1700) / 1620;
	END_IF;

END_FUNCTION

FUNCTION DAY_OF_MONTH:INT
	VAR_INPUT
		IDATE :	UDINT;
	END_VAR

	day_of_month := day_of_year_UDINT(idate);

	IF leap_of_Date(idate) THEN
		CASE day_of_month OF
			32..60	:	day_of_month := day_of_month - 31;
			61..91	:	day_of_month := day_of_month - 60;
			92..121 :	day_of_month := day_of_month - 91;
			122..152:	day_of_month := day_of_month - 121;
			153..182:	day_of_month := day_of_month - 152;
			183..213:	day_of_month := day_of_month - 182;
			214..244:	day_of_month := day_of_month - 213;
			245..274:	day_of_month := day_of_month - 244;
			275..305:	day_of_month := day_of_month - 274;
			306..335:	day_of_month := day_of_month - 305;
			336..366:	day_of_month := day_of_month - 335;
		END_CASE;
	ELSE
		CASE day_of_month OF
			32..59	:	day_of_month := day_of_month - 31;
			60..90	:	day_of_month := day_of_month - 59;
			91..120 :	day_of_month := day_of_month - 90;
			121..151:	day_of_month := day_of_month - 120;
			152..181:	day_of_month := day_of_month - 151;
			182..212:	day_of_month := day_of_month - 181;
			213..243:	day_of_month := day_of_month - 212;
			244..273:	day_of_month := day_of_month - 243;
			274..304:	day_of_month := day_of_month - 273;
			305..334:	day_of_month := day_of_month - 304;
			335..365:	day_of_month := day_of_month - 334;
		END_CASE;
	END_IF;

END_FUNCTION

FUNCTION LEAP_OF_DATE:BOOL

	VAR_INPUT
		IDATE :	UDINT;
	END_VAR

	LEAP_OF_DATE := SHL(UDINT_TO_DWORD((idate + UDINT#43200) / UDINT#31557600), 30) = DWORD#16#80000000;
END_FUNCTION

FUNCTION DAY_OF_YEAR:INT
	VAR_INPUT
		IDATE :	UDINT;
	END_VAR

	DAY_OF_YEAR := UDINT_TO_INT(((idate) / UDINT#86400) MOD UDINT#1461);
	IF DAY_OF_YEAR > 729 THEN
		IF DAY_OF_YEAR > 1095 THEN DAY_OF_YEAR := DAY_OF_YEAR - 1095; ELSE DAY_OF_YEAR := DAY_OF_YEAR - 729; END_IF;
	ELSIF DAY_OF_YEAR > 364 THEN
		DAY_OF_YEAR := DAY_OF_YEAR - 364;
	ELSE
		DAY_OF_YEAR := DAY_OF_YEAR + 1;
	END_IF;
END_FUNCTION

FUNCTION MONTH_OF_DATE:INT

	VAR_INPUT
		IDATE :	UDINT;
	END_VAR

	MONTH_OF_DATE := DAY_OF_YEAR(idate);
	IF MONTH_OF_DATE < 32 THEN
		MONTH_OF_DATE := 1;
	ELSIF LEAP_OF_DATE((IDATE)) THEN
		MONTH_OF_DATE := (MONTH_OF_DATE * 53 + 1668) / 1623;
	ELSE
		MONTH_OF_DATE := (MONTH_OF_DATE * 53 + 1700) / 1620;
	END_IF;
END_FUNCTION

FUNCTION YEAR_OF_DATE:INT
	VAR_INPUT
		IDATE :	UDINT;
	END_VAR

	YEAR_OF_DATE := UDINT_TO_INT((idate+UDINT#43200) / UDINT#31557600 + UDINT#1970);
END_FUNCTION

FUNCTION _INT_TO_UDINT:UDINT
	VAR_INPUT
		IN :	INT;
	END_VAR

	_INT_TO_UDINT := DINT_TO_UDINT(INT_TO_DINT(IN));
END_FUNCTION

FUNCTION DT_TO_DATE:UDINT
	VAR_INPUT
		IN :	UDINT;
	END_VAR

	DT_TO_DATE := (IN / UDINT#86400) * UDINT#86400;
END_FUNCTION

FUNCTION SET_DT:UDINT

	VAR_INPUT
		YEAR : INT;
		MONTH :	INT;
		DAY : INT;
		HOUR : INT;
		MINUTE : INT;
		SECOND : INT;
	END_VAR

	SET_DT := SET_DATE(YEAR, MONTH, DAY) + _INT_TO_UDINT(SECOND) + _INT_TO_UDINT(MINUTE) * UDINT#60 + _INT_TO_UDINT(HOUR) * UDINT#3600;

END_FUNCTION

FUNCTION SET_DATE:UDINT

	VAR_INPUT
		YEAR :	INT;
		MONTH :	INT;
		DAY :	INT;
	END_VAR

	VAR
		count :	INT;
	END_VAR

	IF month > 2 THEN
		count := (month - 1) * 30;
		IF month > 7 THEN
			count := count + DWORD_TO_INT(SHR(DINT_TO_DWORD(INT_TO_DINT(month) - INT_TO_DINT(3)),1));
		ELSE
			count := count + DWORD_TO_INT(SHR(DINT_TO_DWORD(INT_TO_DINT(month) - INT_TO_DINT(4)),1));
		END_IF;
		IF SHL(INT_TO_WORD(year),14) = WORD#0 THEN
			count := count + 1;
		END_IF;
	ELSE
		count := (month - 1) * 31;
	END_IF;
	SET_DATE := (_INT_TO_UDINT(count + day - 1) + DWORD_TO_UDINT(SHR(UDINT_TO_DWORD(_INT_TO_UDINT(year) * UDINT#1461 - UDINT#2878169), 2))) * UDINT#86400;

END_FUNCTION

FUNCTION MONTH_END:UDINT

	VAR_INPUT
		IDATE :	UDINT;
	END_VAR

	MONTH_END := SET_DATE(YEAR_OF_DATE(idate),MONTH_OF_DATE(idate)+1,1) - UDINT#86400;

END_FUNCTION

FUNCTION YEAR_END:UDINT

	VAR_INPUT
		Y :	INT;
	END_VAR

	YEAR_END := DWORD_TO_UDINT(SHR(UDINT_TO_DWORD(INT_TO_UDINT(y) * UDINT#1461 - UDINT#2876712), 2)) * UDINT#86400;

END_FUNCTION

FUNCTION LEAP_DAY:BOOL

	VAR_INPUT
		IDATE :	UDINT;
	END_VAR

	LEAP_DAY := IDATE MOD UDINT#126230400 = UDINT#68169600;

END_FUNCTION

FUNCTION BIT_LOAD_B:BYTE
	VAR_INPUT
		IN :	BYTE;
		VAL :	BOOL;
		POS :	INT;
	END_VAR

	IF VAL THEN
		BIT_LOAD_B := in OR SHL(BYTE#1,pos);
	ELSE
		BIT_LOAD_B := in AND (NOT SHL(BYTE#1,pos));
	END_IF;
END_FUNCTION

FUNCTION BIT_OF_DWORD : BOOL
  VAR_INPUT
    IN : DWORD;
    N : INT;
  END_VAR

  BIT_OF_DWORD := (SHR(in,N) AND 16#00000001) > 0;
END_FUNCTION

FUNCTION_BLOCK TIMER_P4_Block

	VAR_INPUT
		DTIME :	UDINT;
		TREF_0 :	UDINT;
		TREF_1 :	UDINT;
		HOLY :	BOOL;
		L0 :	BOOL;
		L1 :	BOOL;
		L2 :	BOOL;
		L3 :	BOOL;
		OFS :	BYTE;
		ENQ :	BOOL;
		MAN :	BOOL;
		MI :	BYTE;
		RST :	BOOL;
	END_VAR

	VAR_IN_OUT
		PROG :	oscat_TIMER_EVENT;
	END_VAR

	VAR_OUTPUT
		Q0 :	BOOL;
		Q1 :	BOOL;
		Q2 :	BOOL;
		Q3 :	BOOL;
		STATUS :	BYTE;
	END_VAR

	VAR
		day_start :	UDINT;
		start :	UDINT;
		event :	oscat_TIMER_EVENT_DATA;
		pos :	INT;
		last_execute :	UDINT;
		current_day :	DINT;
		mask :	BYTE;
		ma :	oscat_arb_0_3;
		mo :	oscat_arb_0_3;
		qn :	oscat_TP4_qn;
		qs :	oscat_TP4_qn;
		channel :	INT;
		tx :	UDINT;
		array_max :	INT := 63;
		channel_max :	INT := 3;
	END_VAR

	IF RST THEN
		last_execute := UDINT#00;
		FOR pos := 0 TO ARRAY_MAX DO
			IF (PROG[pos].CHANNEL >= OFS) AND (_BYTE_TO_INT(PROG[pos].CHANNEL) < (_BYTE_TO_INT(OFS) + 4)) THEN PROG[pos].LAST := last_execute; END_IF;
		END_FOR;

		FOR pos := 0 TO channel_max DO
			qs[pos] := FALSE;
		END_FOR;

	ELSIF dtime <> last_execute THEN
		last_execute := DTIME;

		day_start := DATE_TO_DT(_DT_TO_DATE_B(DTIME));

		FOR pos := 0 TO channel_max DO qn[pos] := FALSE; END_FOR;

		FOR pos := 0 TO ARRAY_MAX DO
			event := prog[pos];
			channel := _BYTE_TO_INT(event.CHANNEL) - _BYTE_TO_INT(OFS);
			IF (event.TYP > BYTE#0) AND (channel >= 0) AND (channel <= channel_max) THEN
				ma[channel] := event.LAND;
				mo[channel] := event.LOR;
				CASE _BYTE_TO_INT(event.TYP) OF
					1:
						start := day_start + event.start;
						qn[channel] := dtime >= start AND dtime <= start + TIME_TO_UDINT2(event.DURATION);

					2:
						IF (SHR(BYTE#128, DAY_OF_WEEK(_DT_TO_DATE_B(Dtime))) AND event.DAY) > BYTE#0 THEN
							start := day_start + event.start;
							qn[channel] := dtime >= start AND dtime <= start + TIME_TO_UDINT2(event.DURATION);
						END_IF;

					3:
						IF current_day MOD _BYTE_TO_DINT(event.DAY) = DINT#0 THEN
							start := day_start + event.start;
							qn[channel] := dtime >= start AND dtime <= start + TIME_TO_UDINT2(event.DURATION);
						END_IF;

					10:
						IF DAY_OF_WEEK(_DT_TO_DATE_B(DTIME)) = BYTE_TO_INT(event.DAY) THEN
							start := day_start + event.start;
							qn[channel] := dtime >= start AND dtime <= start + TIME_TO_UDINT2(event.DURATION);
						END_IF;

					20:
						IF DAY_OF_MONTH(_DT_TO_DATE_B(DTIME)) = BYTE_TO_INT(event.DAY) THEN
							start := day_start + event.start;
							qn[channel] := dtime >= start AND dtime <= start + TIME_TO_UDINT2(event.DURATION);
						END_IF;

					21:
						IF _DT_TO_DATE_B(DTIME) = MONTH_END(_DT_TO_DATE_B(dtime)) THEN
							start := day_start + event.start;
							qn[channel] := dtime >= start AND dtime <= start + TIME_TO_UDINT2(event.DURATION);
						END_IF;

					30:
						IF DAY_OF_YEAR(_DT_TO_DATE_B(DTIME)) = BYTE_TO_INT(event.DAY) THEN
							start := day_start + event.start;
							qn[channel] := dtime >= start AND dtime <= start + TIME_TO_UDINT2(event.DURATION);
						END_IF;

					31:
						IF _DT_TO_DATE_B(DTIME) = YEAR_END(YEAR_OF_DATE(_DT_TO_DATE_B(dtime))) THEN
							start := day_start + event.start;
							qn[channel] := dtime >= start AND dtime <= start + TIME_TO_UDINT2(event.DURATION);
						END_IF;

					40:
						IF LEAP_DAY(_DT_TO_DATE_B(dtime)) THEN
							start := day_start + event.start;
							qn[channel] := dtime >= start AND dtime <= start + TIME_TO_UDINT2(event.DURATION);
						END_IF;

					41:
						IF HOLY THEN
							start := day_start + event.start;
							qn[channel] := dtime >= start AND dtime <= start + TIME_TO_UDINT2(event.DURATION);
						END_IF;

					42:
						IF (Holy OR (DAY_OF_WEEK(_DT_TO_DATE_B(dtime)) = 6) OR (DAY_OF_WEEK(_DT_TO_DATE_B(dtime)) = 7)) THEN
							start := day_start + event.start;
							qn[channel] := dtime >= start AND dtime <= start + TIME_TO_UDINT2(event.DURATION);
						END_IF;

					43:
						IF DAY_OF_WEEK(_DT_TO_DATE_B(dtime)) < 6 THEN
							start := day_start + event.start;
							qn[channel] := dtime >= start AND dtime <= start + TIME_TO_UDINT2(event.DURATION);
						END_IF;

					50:
						CASE _BYTE_TO_INT(prog[pos].DAY) OF
							0:	tx := tref_0;
							1:	tx := tref_1;
						ELSE
							tx := UDINT#0 ;
						END_CASE;
						start := day_start + tx + event.start;
						qn[channel] := dtime >= start AND dtime <= start + TIME_TO_UDINT2(event.DURATION);

					51:
						CASE _BYTE_TO_INT(prog[pos].DAY) OF
							0:	tx := tref_0;
							1:	tx := tref_1;
						ELSE
							tx := UDINT#0;
						END_CASE;
						start := day_start + tx - event.start;
						qn[channel] := dtime >= start AND dtime <= start + TIME_TO_UDINT2(event.DURATION);

					52 :
						CASE _BYTE_TO_INT(prog[pos].DAY) OF
							0:	tx := tref_0;
							1:	tx := tref_1;
						ELSE
							tx := UDINT#0 ;
						END_CASE;
						start := day_start + tx + event.start;
						IF dtime >= start AND day_start > event.LAST THEN
							qs[channel] := TRUE;
							prog[pos].LAST := day_start;
						END_IF;

					53 :
						CASE _BYTE_TO_INT(prog[pos].DAY) OF
							0:	tx := tref_0;
							1:	tx := tref_1;
						ELSE
							tx := UDINT#0 ;
						END_CASE;
						start := day_start + tx + event.start;
						IF dtime >= start AND day_start > event.LAST THEN
							qs[channel] := FALSE;
							prog[pos].LAST := day_start;
						END_IF;

					54 :
						CASE _BYTE_TO_INT(prog[pos].DAY) OF
							0:	tx := tref_0;
							1:	tx := tref_1;
						ELSE
							tx := UDINT#0 ;
						END_CASE;
						start := day_start + tx - event.start;
						IF dtime >= start AND day_start > event.LAST THEN
							qs[channel] := TRUE;
							prog[pos].LAST := day_start;
						END_IF;

					55 :
						CASE _BYTE_TO_INT(prog[pos].DAY) OF
							0:	tx := tref_0;
							1:	tx := tref_1;
						ELSE
							tx := UDINT#0 ;
						END_CASE;
						start := day_start + tx - event.start;
						IF dtime >= start AND day_start > event.LAST THEN
							qs[channel] := FALSE;
							prog[pos].LAST := day_start;
						END_IF;
				END_CASE;
			END_IF;
		END_FOR;
	END_IF;

	mask := BYTE#255;
	mask:=BIT_LOAD_B(mask,L0,0);
	mask:=BIT_LOAD_B(mask,L1,1);
	mask:=BIT_LOAD_B(mask,L2,2);
	mask:=BIT_LOAD_B(mask,L3,3);

	Q0 := ENQ AND ((qn[0] OR qs[0]) AND ((ma[0] AND mask) = ma[0]) OR ((mo[0] AND mask) > BYTE#0) OR (man AND BIT_OF_DWORD(BYTE_TO_DWORD(MI),0)));
	Q1 := ENQ AND ((qn[1] OR qs[1]) AND ((ma[1] AND mask) = ma[1]) OR ((mo[1] AND mask) > BYTE#1) OR (man AND BIT_OF_DWORD(BYTE_TO_DWORD(MI),1)));
	Q2 := ENQ AND ((qn[2] OR qs[2]) AND ((ma[2] AND mask) = ma[2]) OR ((mo[2] AND mask) > BYTE#2) OR (man AND BIT_OF_DWORD(BYTE_TO_DWORD(MI),2)));
	Q3 := ENQ AND ((qn[3] OR qs[3]) AND ((ma[3] AND mask) = ma[3]) OR ((mo[3] AND mask) > BYTE#3) OR (man AND BIT_OF_DWORD(BYTE_TO_DWORD(MI),3)));

	IF NOT enq THEN
		status := BYTE#100;
	ELSIF man THEN
		status := BYTE#101;
	ELSE
		status := BYTE#102;
	END_IF;

END_FUNCTION_BLOCK

PROGRAM program0
	VAR
		DTIME :	UDINT;
		TREF_0 :	UDINT;
		TREF_1 :	UDINT;
		HOLY :	BOOL;
		L0 :	BOOL;
		L1 :	BOOL;
		L2 :	BOOL;
		L3 :	BOOL;
		OFS :	BYTE;
		ENQ :	BOOL;
		MAN :	BOOL;
		MI :	BYTE;
		RST :	BOOL;
		PROG :	oscat_TIMER_EVENT;
		Q0 :	BOOL;
		Q1 :	BOOL;
		Q2 :	BOOL;
		Q3 :	BOOL;
		STATUS :	BYTE;

		func_block : TIMER_P4_Block;
	END_VAR
	func_block.DTIME := DTIME;
	func_block.TREF_0 := TREF_0;
	func_block.TREF_1 := TREF_1;
	func_block.HOLY := HOLY;
	func_block.L0 := L0;
	func_block.L1 := L1;
	func_block.L2 := L2;
	func_block.L3 := L3;
	func_block.OFS := OFS;
	func_block.ENQ := ENQ;
	func_block.MAN := MAN;
	func_block.MI := MI;
	func_block.RST := RST;
	func_block.PROG := PROG;

	func_block();
	PROG  := func_block.PROG;
	Q0  := func_block.Q0;
	Q1  := func_block.Q1;
	Q2  := func_block.Q2;
	Q3  := func_block.Q3;
	STATUS  := func_block.STATUS;
END_PROGRAM

CONFIGURATION Config0
	RESOURCE Res0 ON PLC
		TASK task0(INTERVAL := T#20ms,PRIORITY := 0);
		PROGRAM instance0 WITH task0 : program0;
	END_RESOURCE
END_CONFIGURATION

(* ---- WORLD_WEATHER.ST ---- *)
TYPE
  oscat_STRING30              : STRING;
  oscat_STRING250             : STRING;
  oscat_STRING8               : STRING;
  oscat_STRING60               : STRING;
  oscat_STRING3               : STRING;
  oscat_STRING10               : STRING;
END_TYPE

TYPE
  oscat_IP_FIFO128_DATA  : ARRAY [1..128] OF BYTE;
  oscat_Mailbox  : ARRAY [1..16] OF BYTE;

  oscat_IP_FIFO_DATA :
  STRUCT
	X       : oscat_IP_FIFO128_DATA; (* IP_ID FIFO Speicher          *)
	Y       : oscat_IP_FIFO128_DATA; (* IP_ID Z�hler                 *)
	ID      : BYTE;                  (* h�chste vergabene id         *)
	MAX_ID  : BYTE;                  (* maximal Anmeldungen pro ID   *)
    INIT    : BOOL;                  (* Initialisierung durchgef�hrt *)
	EMPTY   : BOOL;                  (* FIFO leer                    *)
	FULL    : BOOL;                  (* FIFO voll                    *)
	TOP     : INT;                   (* maximale anzahl in FIFO      *)
	NW      : INT;                   (* Schreibzeiger                *)
	NR      : INT;                   (* Lesezeiger                   *)
  END_STRUCT;

  oscat_IP_C:
  STRUCT
  	C_MODE:			BYTE;          		(*W Mode: TCP/UCP AKTIV/PASSIV                               *)
	C_PORT:         WORD;          		(*W Portnummer                                               *)
	C_IP:           DWORD;         		(*W IP-Adresse gepackt wwxxyyzz = www.xxx.yyy.zzz            *)
    C_STATE:        BYTE;          		(*R Verbindungsstatus ON/OFF + Flanke ON/OFF                 *)
	C_ENABLE:       BOOL;          		(*W Freigabe f�r Connect                                     *)
    R_OBSERVE:      BOOL;          		(*W Empfang ueberwachen                                      *)
    TIME_RESET:     BOOL;          		(*W Alle Timer ruecksetzen                                   *)
	ERROR:          DWORD;         		(*R vvwwxxyy (vv = CON_ERROR, ww = SEN_ERROR, xx = REC_ERROR *)
    FIFO:           oscat_IP_FIFO_DATA; (*I IP FIFO Struktur                                         *)
	MAILBOX:		oscat_Mailbox;		(*I Mailbox: Datenbereich f�r Bausteindatenaustausch         *)
  END_STRUCT;

  oscat_XML_CONTROL:
  STRUCT
    COMMAND:             WORD;            (*W                 *)
    WATCHDOG:            TIME;            (*W                 *)
    START_POS:           UINT;            (*W                 *)
    STOP_POS:            UINT;            (*W                 *)
    COUNT:               UINT;            (*R                 *)
    TYP:                 INT;             (*R                 *)
    LEVEL:               UINT;            (*R                 *)
    PATH:                oscat_STRING250; (*R                 *)
    ELEMENT:             oscat_STRING250; (*R                 *)
    ATTRIBUTE:           oscat_STRING250; (*R                 *)
    VALUE:               oscat_STRING250; (*R                 *)
    BLOCK1_START:        UINT;            (*R                 *)
    BLOCK1_STOP:         UINT;            (*R                 *)
    BLOCK2_START:        UINT;            (*R                 *)
    BLOCK2_STOP:         UINT;            (*R                 *)
  END_STRUCT;

  (* --------- WORLD WEATHER --------- *)

  oscat_WORLD_WEATHER_CUR :
  STRUCT
	OBSERVATION_TIME : oscat_STRING8;
	TEMP_C           : INT;
	WEATHER_CODE     : INT;
	WEATHER_DESC 	 : oscat_STRING60;
	WEATHER_ICON     : INT;
	WIND_SPEED_MILES : INT;
	WIND_SPEED_KMPH  : INT;
	WIND_DIR_DEGREE  : INT;
	WIND_DIR16POINT  : oscat_STRING3;
	PRECIPMM         : REAL;
	HUMIDITY         : INT;
	VISIBILITY       : INT;
	PRESSURE         : INT;
	CLOUDOVER        : INT;
  END_STRUCT;

  oscat_WORLD_WEATHER_DAY :
  STRUCT
	DATE_OF_DAY      : oscat_STRING10;
	TEMP_MAX_C       : INT;
	TEMP_MAX_F       : INT;
	TEMP_MIN_C       : INT;
	TEMP_MIN_F       : INT;
	WIND_SPEED_MILES : INT;
	WIND_SPEED_KMPH  : INT;
	WIND_DIR_DEGREE  : INT;
	WIND_DIR16POINT  : oscat_STRING3;
	WEATHER_CODE     : INT;
	WEATHER_DESC     : oscat_STRING60;
	WEATHER_ICON     : INT;
	PRECIPMM         : REAL;
  END_STRUCT;

  oscat_WORLD_WEATHER_DAY_ARR : ARRAY [0..4] OF oscat_WORLD_WEATHER_DAY;

  oscat_WORLD_WEATHER_DATA :
  STRUCT
	CUR : oscat_WORLD_WEATHER_CUR;
	DAY : oscat_WORLD_WEATHER_DAY_ARR;
  END_STRUCT;

  oscat_WORLD_WEATHER_aI0_41 : ARRAY[0..41] OF INT;

END_TYPE

TYPE
  oscat_NW_BUF_LONG  : ARRAY [0..4095] OF BYTE;

  oscat_NETWORK_BUFFER :
  STRUCT
    SIZE   : UINT;
    BUFFER : oscat_NW_BUF_LONG;
  END_STRUCT;

END_TYPE

FUNCTION_BLOCK WORLD_WEATHER_Block

	VAR_INPUT
		ACTIVATE :	BOOL;
		LATITUDE :	REAL;
		LONGITUDE :	REAL;
		KEY :	oscat_STRING30;
	END_VAR

	VAR_OUTPUT
		BUSY :	BOOL;
		DONE :	BOOL;
		ERROR_C :	DWORD;
		ERROR_T :	BYTE;
	END_VAR

	VAR_IN_OUT
		IP_C :	oscat_IP_C;
		S_BUF :	oscat_NETWORK_BUFFER;
		R_BUF :	oscat_NETWORK_BUFFER;
		WW :	oscat_WORLD_WEATHER_DATA;
	END_VAR

	VAR
		CHK_REAL :	CHK_REAL;
		REAL_TO_STRF :	REAL_TO_STRF;
		URL_DATA :	oscat_url;
		DNS_CLIENT :	DNS_CLIENT;
		HTTP_GET :	HTTP_GET;
		CPB :	CSV_PARSER_BUF;
		STRING_TO_URL :	STRING_TO_URL;
		FLOAT_TO_REAL :	FLOAT_TO_REAL;
		last_state :	BOOL;
		value_int :	INT;
		value_real :	REAL;
		v_real :	REAL;
		state :	INT;
		url_str :	oscat_STRING250;
		offset :	UDINT;
		size :	INT;
		sep :	BYTE;
		cnt :	INT;
		day :	INT;
		idx :	INT;
		run :	BYTE;
		result :	BYTE;
		value :	oscat_STRING250;
		DEC_TO_INT :	DEC_TO_INT;
		pos :	INT;
	END_VAR

	CASE state OF

	00:
		IF ACTIVATE AND NOT last_state THEN
			state := 20;
			DONE := FALSE;
			BUSY := TRUE;
			ERROR_C := DWORD#0;
			ERROR_T := BYTE#0;
		END_IF;

	20:
		REAL_TO_STRF(IN:=LATITUDE,N:=6,D:='.');
		url_str := CONCAT('http://free.worldweatheronline.com/feed/weather.ashx?q=',REAL_TO_STRF.REAL_TO_STRF);
		url_str := CONCAT(url_str,',');
		REAL_TO_STRF(IN:=LONGITUDE,N:=6,D:='.');
		url_str := CONCAT(url_str,REAL_TO_STRF.REAL_TO_STRF);
		url_str := CONCAT(url_str,'&format=csv&num_of_days=5&key=');
		url_str := CONCAT(url_str,key);

		STRING_TO_URL(STR:=url_str, DEFAULT_PROTOCOL:='', DEFAULT_PATH:='' );
		URL_DATA:=STRING_TO_URL.STRING_TO_URL;

		state := 40;

	40:
		IF DNS_CLIENT.DONE THEN
			state := 60;
		ELSIF (DNS_CLIENT.ERROR > DWORD#00) THEN
			ERROR_C := DNS_CLIENT.ERROR;
			ERROR_T := BYTE#01;
			state   := 100;
		END_IF;

	60:
		IF HTTP_GET.DONE THEN
			sep := BYTE#0;
			idx := 0;
			day := 0;
			cnt := 0;
			OFFSET := UINT_TO_UDINT(HTTP_GET.BODY_START);
			size := UINT_TO_INT(HTTP_GET.BODY_STOP);
			run := BYTE#1;
			state := 80;

		ELSIF (HTTP_GET.ERROR > DWORD#00) THEN
			ERROR_C := HTTP_GET.ERROR;
			ERROR_T := BYTE#02;
			state := 100;
		END_IF;

	80:	IF run = BYTE#0 THEN
			run := BYTE#1;
			IF result = BYTE#1 OR result = BYTE#2 THEN
				value_int := 0;
				value_real := 0.0;
				IF LEN(value) <= 20 THEN
					FLOAT_TO_REAL(FLT:=value);
					v_real := FLOAT_TO_REAL.FLOAT_TO_REAL;
					CHK_REAL(X := v_real);
					IF CHK_REAL.CHK_REAL = BYTE#0 THEN
						value_real := v_real;
						value_int := REAL_TO_INT(value_real);
					END_IF;
				END_IF;
				cnt := cnt + 1;
				IF cnt >=8 AND cnt <= 87 THEN
					IF cnt > 22 THEN
						CASE idx OF
						00:	WW.DAY[day].DATE_OF_DAY := value;
						01:	WW.DAY[day].TEMP_MAX_C := value_int;
						02:	WW.DAY[day].TEMP_MAX_F := value_int;
						03:	WW.DAY[day].TEMP_MIN_C := value_int;
						04:	WW.DAY[day].TEMP_MIN_F := value_int;
						05:	WW.DAY[day].WIND_SPEED_MILES := value_int;
						06:	WW.DAY[day].WIND_SPEED_KMPH := value_int;
						07:	WW.DAY[day].WIND_DIR_DEGREE := value_int;
						08:	WW.DAY[day].WIND_DIR16POINT := value;
						09:	WW.DAY[day].WEATHER_CODE := value_int;
						10:	pos := FIND(value, '/wsymbol_');
							IF pos > 0 AND LEN(value) > pos + 13 THEN
								DEC_TO_INT(DEC:=MID(value,4,pos + 9));
								WW.DAY[day].WEATHER_ICON := DEC_TO_INT.DEC_TO_INT;
							ELSE
								WW.DAY[day].WEATHER_ICON := 0;
							END_IF;
						11:	WW.DAY[day].WEATHER_DESC := value;
						12:	WW.DAY[day].PRECIPMM := value_real;
						END_CASE;
						idx := idx + 1;
						IF idx > 12 THEN
							idx := 0;
							day := day + 1;
						END_IF;
					ELSE
						CASE cnt OF
						08:	sep := BYTE#44;
						09:	WW.CUR.OBSERVATION_TIME := value;
						10:	WW.CUR.TEMP_C := value_int;
						11:	WW.CUR.WEATHER_CODE := value_int;
						12:	pos := FIND(value, '/wsymbol_');
							IF pos > 0 AND LEN(value) > pos + 13 THEN
								DEC_TO_INT(DEC:=MID(value,4,pos + 9));
								WW.CUR.WEATHER_ICON := DEC_TO_INT.DEC_TO_INT;
							ELSE
								WW.CUR.WEATHER_ICON := 0;
							END_IF;
						13:	WW.CUR.WEATHER_DESC := value;
						14:	WW.CUR.WIND_SPEED_MILES := value_int;
						15:	WW.CUR.WIND_SPEED_KMPH := value_int;
						16:	WW.CUR.WIND_DIR_DEGREE := value_int;
						17:	WW.CUR.WIND_DIR16POINT := value;
						18:	WW.CUR.PRECIPMM := value_real;
						19:	WW.CUR.HUMIDITY := value_int;
						20:	WW.CUR.VISIBILITY := value_int;
						21:	WW.CUR.PRESSURE := value_int;
						22:	WW.CUR.CLOUDOVER := value_int;
						END_CASE;
					END_IF;
				END_IF;
			ELSIF result = BYTE#10 THEN
				DONE  := TRUE;
				run := BYTE#0;
				state := 100;
			END_IF;
		END_IF;

	100:
		IF (NOT HTTP_GET.DONE) THEN
			state := 0;
			BUSY := FALSE;
			DONE := ERROR_T = BYTE#0;
		END_IF;

	END_CASE;

	DNS_CLIENT.IP_C     := IP_C;
	DNS_CLIENT.S_BUF    := S_BUF;
	DNS_CLIENT.R_BUF    := R_BUF;
	DNS_CLIENT.DOMAIN   := URL_DATA.DOMAIN;
	DNS_CLIENT.IP4_DNS  := DWORD#00;
	DNS_CLIENT.ACTIVATE := state=40;
	DNS_CLIENT();
	IP_C  := DNS_CLIENT.IP_C;
	S_BUF := DNS_CLIENT.S_BUF;
	R_BUF := DNS_CLIENT.R_BUF;

	HTTP_GET.IP_C        := IP_C;
	HTTP_GET.S_BUF       := S_BUF;
	HTTP_GET.R_BUF       := R_BUF;
	HTTP_GET.IP4         := DNS_CLIENT.IP4;
	HTTP_GET.GET         := state=60;
	HTTP_GET.MODE        := BYTE#2;
	HTTP_GET.UNLOCK_BUF  := state=100;
	HTTP_GET.URL_DATA    := URL_DATA;
	HTTP_GET();
	IP_C     := HTTP_GET.IP_C;
	S_BUF    := HTTP_GET.S_BUF;
	R_BUF    := HTTP_GET.R_BUF;
	URL_DATA := HTTP_GET.URL_DATA;

	CPB(SEP:=sep,RUN:=run,OFFSET:=offset,VALUE:=value,PT:=R_BUF);
	run:=CPB.RUN;
	offset:=CPB.OFFSET;
	value:=CPB.VALUE;
	R_BUF:=CPB.PT;
	result:=CPB.RESULT;

	last_state := ACTIVATE;

END_FUNCTION_BLOCK

PROGRAM program0
	VAR
		ACTIVATE :	BOOL;
		LATITUDE :	REAL;
		LONGITUDE :	REAL;
		KEY :	oscat_STRING30;
		IP_C :	oscat_IP_C;
		S_BUF :	oscat_NETWORK_BUFFER;
		R_BUF :	oscat_NETWORK_BUFFER;
		WW :	oscat_WORLD_WEATHER_DATA;
		BUSY :	BOOL;
		DONE :	BOOL;
		ERROR_C :	DWORD;
		ERROR_T :	BYTE;

		func_block : WORLD_WEATHER_Block;
	END_VAR
	func_block.ACTIVATE := ACTIVATE;
	func_block.LATITUDE := LATITUDE;
	func_block.LONGITUDE := LONGITUDE;
	func_block.KEY := KEY;
	func_block.IP_C := IP_C;
	func_block.S_BUF := S_BUF;
	func_block.R_BUF := R_BUF;
	func_block.WW := WW;

	func_block();
	IP_C  := func_block.IP_C;
	S_BUF  := func_block.S_BUF;
	R_BUF  := func_block.R_BUF;
	WW  := func_block.WW;
	BUSY  := func_block.BUSY;
	DONE  := func_block.DONE;
	ERROR_C  := func_block.ERROR_C;
	ERROR_T  := func_block.ERROR_T;
END_PROGRAM

CONFIGURATION Config0
	RESOURCE Res0 ON PLC
		TASK task0(INTERVAL := T#20ms,PRIORITY := 0);
		PROGRAM instance0 WITH task0 : program0;
	END_RESOURCE
END_CONFIGURATION

(* ---- A_TRIG.ST ---- *)
FUNCTION_BLOCK A_TRIG

	VAR_INPUT
		IN :	REAL;
		RES :	REAL;
	END_VAR

	VAR_OUTPUT
		Q :	BOOL;
		D :	REAL;
	END_VAR

	VAR
		last_in :	REAL;
	END_VAR

	D := IN - LAST_IN;
	IF ABS(D) >= res THEN
		Q := TRUE;
		last_in := IN;
	ELSE
		Q := FALSE;
	END_IF;

END_FUNCTION_BLOCK

PROGRAM program0
	VAR
	    LocalVar0 : REAL;
		LocalVar1 : REAL;
		LocalOUT1  : BOOL;
		LocalOUT2  : REAL;
		func_block : A_TRIG;
  	END_VAR
	func_block.IN := LocalVar0;
    func_block.RES := LocalVar1;
	func_block();
	LocalOUT1 := func_block.Q;
	LocalOUT2 := func_block.D;
END_PROGRAM

CONFIGURATION Config0
  	RESOURCE Res0 ON PLC
    	TASK task0(INTERVAL := T#20ms,PRIORITY := 0);
    	PROGRAM instance0 WITH task0 : program0;
  	END_RESOURCE
END_CONFIGURATION

(* ---- ACTUATOR_2P.ST ---- *)
FUNCTION UDINT_TO_TIME2:TIME

	VAR_INPUT
		IN :	UDINT;
	END_VAR

	UDINT_TO_TIME2 := DINT_TO_TIME(UDINT_TO_DINT(IN));

END_FUNCTION

FUNCTION_BLOCK T_PLC_MS_block
	VAR_OUTPUT
		T_PLC_MS :	UDINT;
	END_VAR

	VAR_EXTERNAL
		PLC_TICKS_PER_SEC :	INT;
		PLC_SYS_TICK_CNT :	DINT;
	END_VAR

	VAR
		debug :	BOOL;(*Debug-Mode ON / OFF*)
		N :	INT;(*Debug-Faktor*)
		Offset :	UDINT;(*Debug-Offset*)
		temp :	DWORD := DWORD#1;(*Debug-Offset*)
		mode :	BOOL;(*modus*)
		faktor :	UDINT;(*Systemtakt-Faktor*)
		init :	BOOL;
		v_plc_ticks_per_sec :	UDINT;
		base :	UDINT := UDINT#1000;
	END_VAR

	IF init = FALSE THEN
		v_plc_ticks_per_sec := INT_TO_UDINT(PLC_TICKS_PER_SEC);
		IF v_plc_ticks_per_sec = UDINT#1024 THEN
			faktor := UDINT#1;
			mode := FALSE;
		ELSIF v_plc_ticks_per_sec > UDINT#0 THEN
			IF v_plc_ticks_per_sec <= base THEN
				faktor := base / v_plc_ticks_per_sec;
				mode := FALSE;
			ELSE
				faktor := v_plc_ticks_per_sec / base;
				mode := TRUE;
			END_IF;
		ELSE
			faktor := UDINT#1;
		END_IF;
		init := TRUE;
	END_IF;

	IF mode THEN
		T_PLC_MS := DINT_TO_UDINT(PLC_SYS_TICK_CNT) / faktor;
	ELSE
		T_PLC_MS := DINT_TO_UDINT(PLC_SYS_TICK_CNT) * faktor;
	END_IF;

	IF debug THEN
		T_PLC_MS := (DWORD_TO_UDINT(SHL(UDINT_TO_DWORD(T_PLC_MS),N) OR SHL(temp,N)) - UDINT#1) + Offset;
	END_IF;

END_FUNCTION_BLOCK

FUNCTION TIME_TO_UDINT2:UDINT
	VAR_INPUT
		X :	TIME;
	END_VAR

	TIME_TO_UDINT2 := DINT_TO_UDINT(TIME_TO_DINT(X));
END_FUNCTION

FUNCTION FRMP_B:BYTE
	VAR_INPUT
		START :	BYTE;
		DIR :	BOOL;
		TD :	TIME;
		TR :	TIME;
	END_VAR

	IF TD < TR THEN
		FRMP_B := MIN(UDINT_TO_BYTE(DWORD_TO_UDINT(SHL(TIME_TO_DWORD(TD), 8)) / TIME_TO_UDINT2(TR)), SEL(DIR, START, USINT_TO_BYTE(USINT#255 - BYTE_TO_USINT(START))));
		IF DIR THEN
			FRMP_B := USINT_TO_BYTE(BYTE_TO_USINT(START) + BYTE_TO_USINT(FRMP_B));
		ELSE
			FRMP_B := USINT_TO_BYTE(BYTE_TO_USINT(START) - BYTE_TO_USINT(FRMP_B));
		END_IF;
	ELSE
		FRMP_B := SEL(DIR, BYTE#0, BYTE#255);
	END_IF;
END_FUNCTION

FUNCTION_BLOCK _RMP_B
	VAR_INPUT
		DIR :	BOOL;
		E :	BOOL := TRUE;
		TR :	TIME;
	END_VAR

	VAR_IN_OUT
		RMP :	BYTE;
	END_VAR

	VAR
		T_PLC_MS :	T_PLC_MS_block;
		tx :	TIME;
		tl :	TIME;
		tn :	TIME;
		init :	BOOL;
		last_dir :	BOOL;
		start :	BYTE;
	END_VAR

	T_PLC_MS();
	tx := UDINT_TO_TIME(T_PLC_MS.T_PLC_MS);

	IF E AND init AND (dir = last_dir) AND (RMP <> SEL(DIR, BYTE#0, BYTE#255)) AND TR = tn THEN
		RMP := FRMP_B(start, DIR, tx - tl, TR);
	ELSE
		init := TRUE;
		tl := tx;
		tn := tr;
		start := RMP;
	END_IF;
	last_dir := dir;
END_FUNCTION_BLOCK

FUNCTION_BLOCK AUTORUN_Block

	VAR_INPUT
		IN :	BOOL;
		TEST :	BOOL;
		ARE :	BOOL := TRUE;
		TRUN :	TIME;
		TOFF :	TIME;
	END_VAR

	VAR_OUTPUT
		OUT :	BOOL;
		ARO :	BOOL;
	END_VAR

	VAR_IN_OUT
		ARX :	BOOL;
	END_VAR

	VAR
		timer :	_RMP_B;
		val :	BYTE;
	END_VAR

	IF TOFF > T#0s THEN
		timer(DIR:= OUT, TR := SEL(OUT, TOFF, TRUN), RMP := val);
		val := timer.RMP;
	ELSE
		val := BYTE#255;
	END_IF;

	IF (NOT ARX AND ARE AND val = BYTE#0) OR TEST THEN
		val := BYTE#0;
		ARO := TRUE;
		ARX := TRUE;
	ELSIF val = BYTE#255 AND ARO THEN
		ARO := FALSE;
		ARX := FALSE;
	END_IF;

	out := IN OR ARO;

END_FUNCTION_BLOCK

FUNCTION_BLOCK GEN_PULSE_Block

	VAR_INPUT
		ENQ :	BOOL := TRUE;
		PTH :	TIME;
		PTL :	TIME;
	END_VAR

	VAR_OUTPUT
		Q :	BOOL;
	END_VAR

	VAR
		T_PLC_MS :	T_PLC_MS_block;
		tx :	TIME;
		tn :	TIME;
		init :	BOOL;
	END_VAR

	IF enq THEN
		T_PLC_MS();
		tx:= UDINT_TO_TIME(T_PLC_MS.T_PLC_MS);
		IF NOT init THEN init := TRUE; tn := tx; END_IF;
		IF tx - tn >= SEL(Q, PTL, PTH) THEN
			tn := tn + SEL(Q, PTL, PTH);
			Q := NOT Q;
		END_IF;
	ELSE
		Q := FALSE;
		init := FALSE;
	END_IF;

END_FUNCTION_BLOCK

FUNCTION_BLOCK ACTUATOR_2P_Block

	VAR_INPUT
		IN :	BYTE;
		TEST :	BOOL;
		ARE :	BOOL := TRUE;
		CYCLE_TIME :	TIME;
		SENS :	BYTE;
		SELF_ACT_TIME :	TIME;
		SELF_ACT_PULSE :	TIME;
		SELF_ACT_CYCLES :	INT := 1;
	END_VAR

	VAR_OUTPUT
		OUT :	BOOL;
		ARO :	BOOL;
	END_VAR

	VAR_IN_OUT
		ARX :	BOOL;
	END_VAR

	VAR
		timer :	AUTORUN_Block;
		pwgen :	GEN_PULSE_Block;
	END_VAR

	timer(trun := MUL_T_AI(SELF_ACT_PULSE,2 * SELF_ACT_CYCLES), toff := SELF_ACT_TIME, Test := TEST, ARE := ARE, arx := ARX);
	ARX := timer.ARX;
	ARO := timer.ARO;

	IF aro THEN
		pwgen(PTL := SELF_ACT_PULSE, PTH := SELF_ACT_PULSE);
		out := pwgen.Q;
	ELSIF in < sens THEN
		out := FALSE;
	ELSIF BYTE_TO_USINT(in) > USINT#255 - BYTE_TO_USINT(sens) THEN
		out := TRUE;
	ELSE
		pwgen.PTH := (CYCLE_TIME * BYTE_TO_TIME2(BAND_B(IN,SENS))  ) / BYTE_TO_TIME2(BYTE#255);
		pwgen.PTL := CYCLE_TIME - pwgen.PTH;
		pwgen();
		out := pwgen.Q;
	END_IF;

END_FUNCTION_BLOCK

PROGRAM program0
	VAR
		IN :	BYTE;
		TEST :	BOOL;
		ARE :	BOOL := TRUE;
		CYCLE_TIME :	TIME;
		SENS :	BYTE;
		SELF_ACT_TIME :	TIME;
		SELF_ACT_PULSE :	TIME;
		SELF_ACT_CYCLES :	INT := 1;
		OUT :	BOOL;
		ARO :	BOOL;
		func_block : ACTUATOR_2P_Block;
	END_VAR
	func_block.IN := IN;
	func_block.TEST := TEST;
	func_block.ARE := ARE ;
	func_block.CYCLE_TIME := CYCLE_TIME;
	func_block.SENS := SENS;
	func_block.SELF_ACT_TIME := SELF_ACT_TIME ;
	func_block.SELF_ACT_PULSE := SELF_ACT_PULSE;
	func_block.SELF_ACT_CYCLES := SELF_ACT_CYCLES;
	func_block();
	OUT  := func_block.OUT;
	ARO  := func_block.ARO;
END_PROGRAM

CONFIGURATION Config0
	VAR_GLOBAL
		PLC_TICKS_PER_SEC :	INT;
		PLC_SYS_TICK_CNT :	DINT;
	END_VAR
  	RESOURCE Res0 ON PLC
    	TASK task0(INTERVAL := T#20ms,PRIORITY := 0);
    	PROGRAM instance0 WITH task0 : program0;
  	END_RESOURCE
END_CONFIGURATION

(* ---- ACTUATOR_3P.ST ---- *)
FUNCTION UDINT_TO_TIME2:TIME

	VAR_INPUT
		IN :	UDINT;
	END_VAR

	UDINT_TO_TIME2 := DINT_TO_TIME(UDINT_TO_DINT(IN));

END_FUNCTION

FUNCTION_BLOCK T_PLC_MS_block
	VAR_OUTPUT
		T_PLC_MS :	UDINT;
	END_VAR

	VAR_EXTERNAL
		PLC_TICKS_PER_SEC :	INT;
		PLC_SYS_TICK_CNT :	DINT;
	END_VAR

	VAR
		debug :	BOOL;(*Debug-Mode ON / OFF*)
		N :	INT;(*Debug-Faktor*)
		Offset :	UDINT;(*Debug-Offset*)
		temp :	DWORD := DWORD#1;(*Debug-Offset*)
		mode :	BOOL;(*modus*)
		faktor :	UDINT;(*Systemtakt-Faktor*)
		init :	BOOL;
		v_plc_ticks_per_sec :	UDINT;
		base :	UDINT := UDINT#1000;
	END_VAR

	IF init = FALSE THEN
		v_plc_ticks_per_sec := INT_TO_UDINT(PLC_TICKS_PER_SEC);
		IF v_plc_ticks_per_sec = UDINT#1024 THEN
			faktor := UDINT#1;
			mode := FALSE;
		ELSIF v_plc_ticks_per_sec > UDINT#0 THEN
			IF v_plc_ticks_per_sec <= base THEN
				faktor := base / v_plc_ticks_per_sec;
				mode := FALSE;
			ELSE
				faktor := v_plc_ticks_per_sec / base;
				mode := TRUE;
			END_IF;
		ELSE
			faktor := UDINT#1;
		END_IF;
		init := TRUE;
	END_IF;

	IF mode THEN
		T_PLC_MS := DINT_TO_UDINT(PLC_SYS_TICK_CNT) / faktor;
	ELSE
		T_PLC_MS := DINT_TO_UDINT(PLC_SYS_TICK_CNT) * faktor;
	END_IF;

	IF debug THEN
		T_PLC_MS := (DWORD_TO_UDINT(SHL(UDINT_TO_DWORD(T_PLC_MS),N) OR SHL(temp,N)) - UDINT#1) + Offset;
	END_IF;
END_FUNCTION_BLOCK

FUNCTION TIME_TO_UDINT2:UDINT
	VAR_INPUT
		X :	TIME;
	END_VAR

	TIME_TO_UDINT2 := DINT_TO_UDINT(TIME_TO_DINT(X));
END_FUNCTION

FUNCTION FRMP_B:BYTE
	VAR_INPUT
		START :	BYTE;
		DIR :	BOOL;
		TD :	TIME;
		TR :	TIME;
	END_VAR

	IF TD < TR THEN
		FRMP_B := MIN(UDINT_TO_BYTE(DWORD_TO_UDINT(SHL(TIME_TO_DWORD(TD), 8)) / TIME_TO_UDINT2(TR)), SEL(DIR, START, USINT_TO_BYTE(USINT#255 - BYTE_TO_USINT(START))));
		IF DIR THEN
			FRMP_B := USINT_TO_BYTE(BYTE_TO_USINT(START) + BYTE_TO_USINT(FRMP_B));
		ELSE
			FRMP_B := USINT_TO_BYTE(BYTE_TO_USINT(START) - BYTE_TO_USINT(FRMP_B));
		END_IF;
	ELSE
		FRMP_B := SEL(DIR, BYTE#0, BYTE#255);
	END_IF;
END_FUNCTION

FUNCTION_BLOCK _RMP_B
	VAR_INPUT
		DIR :	BOOL;
		E :	BOOL := TRUE;
		TR :	TIME;
	END_VAR

	VAR_IN_OUT
		RMP :	BYTE;
	END_VAR

	VAR
		T_PLC_MS :	T_PLC_MS_block;
		tx :	TIME;
		tl :	TIME;
		tn :	TIME;
		init :	BOOL;
		last_dir :	BOOL;
		start :	BYTE;
	END_VAR

	T_PLC_MS();
	tx := UDINT_TO_TIME(T_PLC_MS.T_PLC_MS);

	IF E AND init AND (dir = last_dir) AND (RMP <> SEL(DIR, BYTE#0, BYTE#255)) AND TR = tn THEN
		RMP := FRMP_B(start, DIR, tx - tl, TR);
	ELSE
		init := TRUE;
		tl := tx;
		tn := tr;
		start := RMP;
	END_IF;
	last_dir := dir;
END_FUNCTION_BLOCK

FUNCTION_BLOCK TREND_DW
	VAR_INPUT
		X :	DWORD;
	END_VAR
	VAR_OUTPUT
		Q :	BOOL;
		TU :	BOOL;
		TD :	BOOL;
		D :	DWORD;
	END_VAR

	VAR
		LAST_X :	DWORD;
	END_VAR

	IF X > last_X THEN
		TU := TRUE;
		TD := FALSE;
		D := UDINT_TO_DWORD(DWORD_TO_UDINT(X) - DWORD_TO_UDINT(last_X));
		Q := TRUE;
	ELSIF X < last_X THEN
		TD := TRUE;
		TU := FALSE;
		D := UDINT_TO_DWORD(DWORD_TO_UDINT(last_X) - DWORD_TO_UDINT(X));
		Q := FALSE;
	ELSE
		TU := FALSE;
		TD := FALSE;
		D := DWORD#0;
	END_IF;
	last_X := X;
END_FUNCTION_BLOCK

FUNCTION_BLOCK _RMP_NEXT_Block
	VAR_INPUT
		E :	BOOL := TRUE;
		IN :	BYTE;
		TR :	TIME;
		TF :	TIME;
		TL :	TIME;
	END_VAR

	VAR_OUTPUT
		DIR :	BOOL;
		UP :	BOOL;
		DN :	BOOL;
	END_VAR

	VAR_IN_OUT
		OUT :	BYTE;
	END_VAR
	VAR
		rmx :	_RMP_B;
		dirx :	TREND_DW;
		t_lock :	TP;
		xen :	BOOL;
		xdir :	BOOL;
	END_VAR

	dirx(X := BYTE_TO_DWORD(in));

	t_lock(in := FALSE, pt := TL);

	IF dirx.TU AND (OUT < IN) THEN
		IF NOT xdir AND xen THEN t_lock(in := TRUE); END_IF;
		xen := TRUE;
		xdir := TRUE;
	ELSIF dirx.TD AND (OUT > IN) THEN
		IF xdir AND xen THEN t_lock(in := TRUE); END_IF;
		xen := TRUE;
		xdir := FALSE;
	ELSIF xen THEN
		IF (xdir AND (out >= in)) OR (NOT xdir AND (out <= in)) THEN
			xen := FALSE;
			IF tl > t#0s THEN t_lock(IN := TRUE); END_IF;
		END_IF;
	END_IF;

	IF NOT t_lock.Q AND xen THEN
		UP := XDIR;
		DIR := XDIR;
		DN := NOT XDIR;
	ELSE
		UP := FALSE;
		DN := FALSE;
	END_IF;

	rmx(rmp := OUT, E := E AND (UP OR DN) , dir := DIR, tr := SEL(dir, TF, TR));
	OUT := rmx.RMP;
END_FUNCTION_BLOCK

FUNCTION _BYTE_TO_INT:INT
	VAR_INPUT
		IN :	BYTE;
	END_VAR

	_BYTE_TO_INT := USINT_TO_INT(BYTE_TO_USINT(IN));
END_FUNCTION

FUNCTION_BLOCK ACTUATOR_3P_Block

	VAR_INPUT
		IN :	BYTE;
		TEST :	BOOL;
		ARE :	BOOL := TRUE;
		END_POS :	BOOL;
		T_RUN :	TIME := T#60s;
		T_EXT :	TIME := T#10s;
		T_CAL :	TIME := T#600s;
		T_DIAG :	TIME := T#10d;
		SWITCH_AVAIL :	BOOL;
	END_VAR

	VAR_OUTPUT
		OUT1 :	BOOL;
		OUT2 :	BOOL;
		POS :	BYTE;
		ERROR :	BOOL;
		STATUS :	BYTE;
	END_VAR

	VAR_IN_OUT
		ARX :	BOOL;
	END_VAR

	VAR
		tx :	TIME;
		_ramp :	_RMP_NEXT_Block;
		next_cal :	TIME;
		next_diag :	TIME;
		last :	TIME;
		start :	TIME;
		T_PLC_MS :	T_PLC_MS_Block;
	END_VAR

	T_PLC_MS();
	tx := UDINT_TO_TIME(T_PLC_MS.T_PLC_MS);

	IF TEST THEN
		status := BYTE#103;
		start := tx;
		ARX := TRUE;
	END_IF;

	CASE _BYTE_TO_INT(status) OF
		0:
			IF ARE AND NOT ARX THEN
				status := BYTE#103;
				start := tx;
				ARX := TRUE;
			END_IF;

		100:
			IF T_DIAG > T#0s AND tx > next_diag AND ARE AND NOT ARX THEN
					status := BYTE#103;
					start := tx;
					ARX := TRUE;

			ELSIF T_CAL > T#0s AND tx > next_cal AND ARE AND NOT ARX THEN
				IF pos > BYTE#127 THEN
					OUT1 := TRUE;
					OUT2 := FALSE;
					_ramp.IN := BYTE#255;
					ARX := TRUE;
				ELSE
					OUT1 := FALSE;
					OUT2 := TRUE;
					_ramp.IN := BYTE#0;
					ARX := TRUE;
				END_IF;
				status := BYTE#101;
				start := tx;
			ELSE
				IF NOT(OUT1 OR OUT2) THEN next_cal := next_cal + (tx-last); END_IF;
				_ramp.IN := IN;
			END_IF;

		101:
			IF tx - start < T_EXT THEN
				next_cal := tx + T_CAL;
			ELSIF SWITCH_AVAIL AND END_POS THEN
				STATUS := BYTE#100;
				ARX := FALSE;
			ELSIF tx - start > T_EXT + T_RUN THEN
				ERROR := SWITCH_AVAIL;
				ARX := FALSE;
			END_IF;

		103:
			IF tx - start < T_EXT THEN
				ERROR := FALSE;
				_ramp.TR := T_RUN;
				_ramp.TF := T_RUN;
				OUT1 := TRUE;
				OUT2 := FALSE;
				_ramp.IN := BYTE#255;
			ELSIF SWITCH_AVAIL AND END_POS THEN
				_ramp.TR := tx - start;
				STATUS := BYTE#104;
			ELSIF tx - start > T_EXT + T_RUN THEN
				ERROR := SWITCH_AVAIL;
				STATUS := BYTE#104;
				start := tx;
			END_IF;

		104:
			IF tx - start < T_ext THEN
				OUT1 := FALSE;
				OUT2 := TRUE;
				_ramp.IN := BYTE#0;
				next_diag := tx + T_DIAG;
			ELSIF SWITCH_AVAIL AND END_POS THEN
				_ramp.TR := tx - start;
				IF DINT_TO_TIME(ABS(TIME_TO_DINT(_ramp.TR) - TIME_TO_DINT(_ramp.TF)) * DINT#10) > T_RUN THEN error := TRUE; END_IF;
				STATUS := BYTE#100;
				ARX := FALSE;
				next_cal := tx + T_CAL;
			ELSIF tx - start > T_EXT + T_RUN THEN
				IF SWITCH_AVAIL THEN ERROR := TRUE; END_IF;
				STATUS := BYTE#100;
				ARX := FALSE;
				next_CAL := tx + T_CAL;
			END_IF;
	END_CASE;

	_ramp(OUT := POS);
	POS := _ramp.OUT;
	IF STATUS = BYTE#100 THEN
		OUT1 := _ramp.UP;
		OUT2 := _ramp.DN;
	END_IF;

	IF SWITCH_AVAIL AND END_POS THEN
		POS := SEL_BYTE(POS > BYTE#127, BYTE#0, BYTE#255);
		next_cal := tx + T_CAL;
	END_IF;

	last := tx;

END_FUNCTION_BLOCK

PROGRAM program0
	VAR
		IN :	BYTE;
		TEST :	BOOL;
		ARE :	BOOL := TRUE;
		END_POS :	BOOL;
		T_RUN :	TIME := T#60s;
		T_EXT :	TIME := T#10s;
		T_CAL :	TIME := T#600s;
		T_DIAG :	TIME := T#10d;
		SWITCH_AVAIL :	BOOL;
		OUT1 :	BOOL;
		OUT2 :	BOOL;
		POS :	BYTE;
		ERROR :	BOOL;
		STATUS :	BYTE;
		func_block : ACTUATOR_3P_Block;
	END_VAR
	func_block.IN := IN;
	func_block.TEST := TEST;
	func_block.ARE := ARE ;
	func_block.END_POS := END_POS;
	func_block.T_RUN := T_RUN;
	func_block.T_EXT := T_EXT;
	func_block.T_CAL := T_CAL ;
	func_block.T_DIAG := T_DIAG;
	func_block.SWITCH_AVAIL := SWITCH_AVAIL;
	func_block();
	OUT1  := func_block.OUT1;
	OUT2  := func_block.OUT2;
	POS  := func_block.POS;
	ERROR  := func_block.ERROR;
	STATUS  := func_block.STATUS;
END_PROGRAM

CONFIGURATION Config0
	VAR_GLOBAL
		PLC_TICKS_PER_SEC :	INT;
		PLC_SYS_TICK_CNT :	DINT;
	END_VAR
  	RESOURCE Res0 ON PLC
    	TASK task0(INTERVAL := T#20ms,PRIORITY := 0);
    	PROGRAM instance0 WITH task0 : program0;
  	END_RESOURCE
END_CONFIGURATION

(* ---- ACTUATOR_A.ST ---- *)
FUNCTION_BLOCK T_PLC_MS_block
	VAR_OUTPUT
		T_PLC_MS :	UDINT;
	END_VAR

	VAR_EXTERNAL
		PLC_TICKS_PER_SEC :	INT;
		PLC_SYS_TICK_CNT :	DINT;
	END_VAR

	VAR
		debug :	BOOL;(*Debug-Mode ON / OFF*)
		N :	INT;(*Debug-Faktor*)
		Offset :	UDINT;(*Debug-Offset*)
		temp :	DWORD := DWORD#1;(*Debug-Offset*)
		mode :	BOOL;(*modus*)
		faktor :	UDINT;(*Systemtakt-Faktor*)
		init :	BOOL;
		v_plc_ticks_per_sec :	UDINT;
		base :	UDINT := UDINT#1000;
	END_VAR

	IF init = FALSE THEN
		v_plc_ticks_per_sec := INT_TO_UDINT(PLC_TICKS_PER_SEC);
		IF v_plc_ticks_per_sec = UDINT#1024 THEN
			faktor := UDINT#1;
			mode := FALSE;
		ELSIF v_plc_ticks_per_sec > UDINT#0 THEN
			IF v_plc_ticks_per_sec <= base THEN
				faktor := base / v_plc_ticks_per_sec;
				mode := FALSE;
			ELSE
				faktor := v_plc_ticks_per_sec / base;
				mode := TRUE;
			END_IF;
		ELSE
			faktor := UDINT#1;
		END_IF;
		init := TRUE;
	END_IF;

	IF mode THEN
		T_PLC_MS := DINT_TO_UDINT(PLC_SYS_TICK_CNT) / faktor;
	ELSE
		T_PLC_MS := DINT_TO_UDINT(PLC_SYS_TICK_CNT) * faktor;
	END_IF;

	IF debug THEN
		T_PLC_MS := (DWORD_TO_UDINT(SHL(UDINT_TO_DWORD(T_PLC_MS),N) OR SHL(temp,N)) - UDINT#1) + Offset;
	END_IF;

END_FUNCTION_BLOCK

FUNCTION_BLOCK CYCLE_4

	VAR_INPUT
		E :	BOOL := TRUE;
		T0 :	TIME;
		T1 :	TIME;
		T2 :	TIME;
		T3 :	TIME;
		S0 :	BOOL;
		SX :	INT;
		SL :	BOOL;
	END_VAR

	VAR_OUTPUT
		STATE :	INT;
	END_VAR

	VAR
		tx :	TIME;
		last :	TIME;
		init :	BOOL;
		T_PLC_MS :	T_PLC_MS_block;
	END_VAR

	T_PLC_MS();
	tx:= UDINT_TO_TIME(T_PLC_MS.T_PLC_MS);

	(* init on first cycle *)
	IF NOT init THEN
		init := TRUE;
		last := tx;
	END_IF;

	IF E THEN
		IF SL THEN
			(* when sx > 0 then the state sx is forced to start *)
			state:= LIMIT(0,SX,3);
			last := tx;
			(* this is to avoid to reset sx from the calling programm it does work fine on codesys but i am not sure about other systems, because we are writing to an input *)
			SL := FALSE;
		ELSE
			CASE state OF
				0 :	(* wait for T0 and switch to next cycle *)
					IF tx - last >= T0 THEN
						state := 1;
						last := tx;
					END_IF;
				1 : (* wait for T1 over 1st cycle *)
					IF tx - last >= T1 THEN
						state := 2;
						last := tx;
					END_IF;
				2 : (* wait for T1 over 1st cycle *)
					IF tx - last >= T2 THEN
						state := 3;
						last := tx;
					END_IF;
				3 : (* wait for T2 over 2nd cycle *)
					IF tx - last >= T3 THEN
						IF S0 THEN State := 0; END_IF; (* if S0 is false, the sequence stops at state 3 *)
						last := tx;
					END_IF;
			END_CASE;
		END_IF;
	ELSE
		state := 0;
		last := tx;
	END_IF;

END_FUNCTION_BLOCK

FUNCTION_BLOCK ACTUATOR_A_Block

	VAR_INPUT
		I1 :	BYTE;
		IS :	BOOL;
		I2 :	BYTE;
		RV :	BOOL;
		DX :	BOOL;
		RUNTIME :	TIME;
		SELF_ACT_TIME :	TIME;
		OUT_MIN :	DWORD;
		OUT_MAX :	DWORD;
	END_VAR

	VAR_OUTPUT
		Y :	DWORD;
	END_VAR

	VAR
		timer :	CYCLE_4;
		dx_edge :	BOOL;
	END_VAR

	timer(T0 := RUNTIME, T1 := RUNTIME, T3 := SELF_ACT_TIME, sl := DX AND NOT dx_edge, sx := 0, S0 := SELF_ACT_TIME > t#0s);
	dx_edge := dx;

	CASE timer.STATE OF
		0:
			Y := OUT_MIN;
		1:
			Y := OUT_MAX;
		3:
			IF rv THEN
				Y := UDINT_TO_DWORD(DWORD_TO_UDINT(OUT_MAX) - (DWORD_TO_UDINT(OUT_MAX) - DWORD_TO_UDINT(OUT_MIN)) * BYTE_TO_UDINT(SEL(IS, I1, I2)) / UDINT#255);
			ELSE
				Y := UDINT_TO_DWORD((DWORD_TO_UDINT(OUT_MAX) - DWORD_TO_UDINT(OUT_MIN)) * BYTE_TO_UDINT(SEL(IS, I1, I2)) / UDINT#255 + DWORD_TO_UDINT(OUT_MIN));
			END_IF;
	END_CASE;

END_FUNCTION_BLOCK

PROGRAM program0
	VAR
		I1 :	BYTE;
		IS :	BOOL;
		I2 :	BYTE;
		RV :	BOOL;
		DX :	BOOL;
		RUNTIME :	TIME;
		SELF_ACT_TIME :	TIME;
		OUT_MIN :	DWORD;
		OUT_MAX :	DWORD;
		Y :	DWORD;
		func_block : ACTUATOR_A_Block;
	END_VAR
	func_block.I1 := I1;
	func_block.IS := IS;
	func_block.I2 := I2 ;
	func_block.RV := RV;
	func_block.DX := DX;
	func_block.RUNTIME := RUNTIME;
	func_block.SELF_ACT_TIME := SELF_ACT_TIME ;
	func_block.OUT_MIN := OUT_MIN;
	func_block.OUT_MAX := OUT_MAX;
	func_block();
	Y  := func_block.Y;
END_PROGRAM

CONFIGURATION Config0
	VAR_GLOBAL
		PLC_TICKS_PER_SEC :	INT;
		PLC_SYS_TICK_CNT :	DINT;
	END_VAR
  	RESOURCE Res0 ON PLC
    	TASK task0(INTERVAL := T#20ms,PRIORITY := 0);
    	PROGRAM instance0 WITH task0 : program0;
  	END_RESOURCE
END_CONFIGURATION

(* ---- ACTUATOR_COIL.ST ---- *)
FUNCTION UDINT_TO_TIME2:TIME

	VAR_INPUT
		IN :	UDINT;
	END_VAR

	UDINT_TO_TIME2 := DINT_TO_TIME(UDINT_TO_DINT(IN));

END_FUNCTION

FUNCTION_BLOCK T_PLC_MS_block
	VAR_OUTPUT
		T_PLC_MS :	UDINT;
	END_VAR

	VAR_EXTERNAL
		PLC_TICKS_PER_SEC :	INT;
		PLC_SYS_TICK_CNT :	DINT;
	END_VAR

	VAR
		debug :	BOOL;(*Debug-Mode ON / OFF*)
		N :	INT;(*Debug-Faktor*)
		Offset :	UDINT;(*Debug-Offset*)
		temp :	DWORD := DWORD#1;(*Debug-Offset*)
		mode :	BOOL;(*modus*)
		faktor :	UDINT;(*Systemtakt-Faktor*)
		init :	BOOL;
		v_plc_ticks_per_sec :	UDINT;
		base :	UDINT := UDINT#1000;
	END_VAR

	IF init = FALSE THEN
		v_plc_ticks_per_sec := INT_TO_UDINT(PLC_TICKS_PER_SEC);
		IF v_plc_ticks_per_sec = UDINT#1024 THEN
			faktor := UDINT#1;
			mode := FALSE;
		ELSIF v_plc_ticks_per_sec > UDINT#0 THEN
			IF v_plc_ticks_per_sec <= base THEN
				faktor := base / v_plc_ticks_per_sec;
				mode := FALSE;
			ELSE
				faktor := v_plc_ticks_per_sec / base;
				mode := TRUE;
			END_IF;
		ELSE
			faktor := UDINT#1;
		END_IF;
		init := TRUE;
	END_IF;

	IF mode THEN
		T_PLC_MS := DINT_TO_UDINT(PLC_SYS_TICK_CNT) / faktor;
	ELSE
		T_PLC_MS := DINT_TO_UDINT(PLC_SYS_TICK_CNT) * faktor;
	END_IF;

	IF debug THEN
		T_PLC_MS := (DWORD_TO_UDINT(SHL(UDINT_TO_DWORD(T_PLC_MS),N) OR SHL(temp,N)) - UDINT#1) + Offset;
	END_IF;
END_FUNCTION_BLOCK

FUNCTION TIME_TO_UDINT2:UDINT
	VAR_INPUT
		X :	TIME;
	END_VAR

	TIME_TO_UDINT2 := DINT_TO_UDINT(TIME_TO_DINT(X));
END_FUNCTION

FUNCTION_BLOCK ACTUATOR_COIL_Block

	VAR_INPUT
		IN :	BOOL;
		SELF_ACT_CYCLE :	TIME := T#10d;
		SELF_ACT_TIME :	TIME := T#1s;
	END_VAR

	VAR_OUTPUT
		OUT :	BOOL;
		STATUS :	BYTE;
	END_VAR

	VAR
		last :	UDINT;
		init :	BOOL;
		tx :	UDINT;
		now :	UDINT;
		T_PLC_MS :	T_PLC_MS_Block;
	END_VAR

	T_PLC_MS();
	now := T_PLC_MS.T_PLC_MS;

	IF NOT init THEN
		last := now;
		init := TRUE;
	ELSIF IN THEN
		OUT := TRUE;
		STATUS := BYTE#101;
		LAST := now;
	ELSE
		OUT := FALSE;
		STATUS := BYTE#100;
		tx := now - last;
		IF (self_act_cycle > T#0s) AND (tx >= TIME_TO_UDINT2(self_act_cycle)) THEN
			OUT := TRUE;
			STATUS := BYTE#102;
			IF tx >= TIME_TO_UDINT2(self_act_cycle + self_act_time) THEN
				last := now;
				OUT := FALSE;
				STATUS := BYTE#100;
			END_IF;
		END_IF;
	END_IF;

END_FUNCTION_BLOCK

PROGRAM program0
	VAR
		IN :	BOOL;
		SELF_ACT_CYCLE :	TIME := T#10d;
		SELF_ACT_TIME :	TIME := T#1s;
		OUT :	BOOL;
		STATUS :	BYTE;
		func_block : ACTUATOR_COIL_Block;
	END_VAR
	func_block.IN := IN;
	func_block.SELF_ACT_CYCLE := SELF_ACT_CYCLE;
	func_block.SELF_ACT_TIME := SELF_ACT_TIME ;
	func_block();
	OUT  := func_block.OUT;
	STATUS  := func_block.STATUS;
END_PROGRAM

CONFIGURATION Config0
	VAR_GLOBAL
		PLC_TICKS_PER_SEC :	INT;
		PLC_SYS_TICK_CNT :	DINT;
	END_VAR
  	RESOURCE Res0 ON PLC
    	TASK task0(INTERVAL := T#20ms,PRIORITY := 0);
    	PROGRAM instance0 WITH task0 : program0;
  	END_RESOURCE
END_CONFIGURATION

(* ---- ACTUATOR_PUMP.ST ---- *)
FUNCTION_BLOCK T_PLC_MS_block
	VAR_OUTPUT
		T_PLC_MS :	UDINT;
	END_VAR

	VAR_EXTERNAL
		PLC_TICKS_PER_SEC :	INT;
		PLC_SYS_TICK_CNT :	DINT;
	END_VAR

	VAR
		debug :	BOOL;(*Debug-Mode ON / OFF*)
		N :	INT;(*Debug-Faktor*)
		Offset :	UDINT;(*Debug-Offset*)
		temp :	DWORD := DWORD#1;(*Debug-Offset*)
		mode :	BOOL;(*modus*)
		faktor :	UDINT;(*Systemtakt-Faktor*)
		init :	BOOL;
		v_plc_ticks_per_sec :	UDINT;
		base :	UDINT := UDINT#1000;
	END_VAR

	IF init = FALSE THEN
		v_plc_ticks_per_sec := INT_TO_UDINT(PLC_TICKS_PER_SEC);
		IF v_plc_ticks_per_sec = UDINT#1024 THEN
			faktor := UDINT#1;
			mode := FALSE;
		ELSIF v_plc_ticks_per_sec > UDINT#0 THEN
			IF v_plc_ticks_per_sec <= base THEN
				faktor := base / v_plc_ticks_per_sec;
				mode := FALSE;
			ELSE
				faktor := v_plc_ticks_per_sec / base;
				mode := TRUE;
			END_IF;
		ELSE
			faktor := UDINT#1;
		END_IF;
		init := TRUE;
	END_IF;

	IF mode THEN
		T_PLC_MS := DINT_TO_UDINT(PLC_SYS_TICK_CNT) / faktor;
	ELSE
		T_PLC_MS := DINT_TO_UDINT(PLC_SYS_TICK_CNT) * faktor;
	END_IF;

	IF debug THEN
		T_PLC_MS := (DWORD_TO_UDINT(SHL(UDINT_TO_DWORD(T_PLC_MS),N) OR SHL(temp,N)) - UDINT#1) + Offset;
	END_IF;

END_FUNCTION_BLOCK

FUNCTION_BLOCK ONTIME_Block

	VAR_INPUT
		IN :	BOOL;
		RST :	BOOL;
	END_VAR

	VAR_IN_OUT
		SECONDS :	UDINT;
		CYCLES :	UDINT;
	END_VAR

	VAR
		tx :	UDINT;
		last :	UDINT;
		edge :	BOOL;
		init :	BOOL;
		ms :	UDINT;
		T_PLC_MS :	T_PLC_MS_Block;
	END_VAR

	T_PLC_MS();
	tx:= T_PLC_MS.T_PLC_MS;

	IF NOT init THEN
		init := TRUE;
		last := tx;
		ms := UDINT#0;
	END_IF;
	IF RST THEN
		SECONDS := UDINT#0;
		CYCLES := UDINT#0;
		last := tx;
		ms := UDINT#0;
	ELSIF IN THEN
		(* add the current milliseconds *)
		ms := (tx - last) + ms;
		IF ms >= UDINT#1000 THEN
			seconds := seconds + UDINT#1;
			ms := ms - UDINT#1000;
		END_IF;
		cycles := cycles + BOOL_TO_UDINT(NOT edge);
	END_IF;
	last := tx;
	edge := in;

END_FUNCTION_BLOCK

FUNCTION_BLOCK ACTUATOR_PUMP_Block

	VAR_INPUT
		IN :	BOOL;
		MANUAL :	BOOL;
		RST :	BOOL := FALSE;
		MIN_ONTIME :	TIME := T#10s;
		MIN_OFFTIME :	TIME := T#10s;
		RUN_EVERY :	TIME := T#10000m;
	END_VAR

	VAR_OUTPUT
		PUMP :	BOOL;
		RUNTIME :	UDINT;
		CYCLES :	UDINT;
	END_VAR

	VAR
		tx :	TIME;
		last_change :	TIME;
		meter :	ONTIME_Block;
		old_man :	BOOL;
		init :	BOOL;
		T_PLC_MS :	T_PLC_MS_Block;
	END_VAR

	T_PLC_MS();
	tx:= UDINT_TO_TIME(T_PLC_MS.T_PLC_MS);

	IF NOT init THEN
		init := TRUE;
		last_change := tx;
	ELSIF rst THEN
		rst := FALSE;
		runtime := UDINT#0;
		cycles := UDINT#0;
	ELSIF manual AND NOT pump AND NOT old_man THEN
		last_change := tx;
		pump := TRUE;
	ELSIF NOT manual AND old_man AND pump AND NOT in THEN
		last_change := tx;
		pump := FALSE;
	ELSIF in AND NOT pump AND tx - last_change >= min_offtime THEN
		last_change := tx;
		pump := TRUE;
	ELSIF pump AND NOT in AND NOT manual AND tx - last_change >= min_ontime THEN
		last_change := tx;
		pump := FALSE;
	ELSIF NOT pump AND (tx - last_change >= run_every) AND (run_every > T#0s) THEN
		last_change := tx;
		pump := TRUE;
	END_IF;

	meter(in := pump, SECONDS := runtime, CYCLES := cycles);
	cycles := meter.CYCLES;
	runtime := meter.SECONDS;

	old_man := manual;

END_FUNCTION_BLOCK

PROGRAM program0
	VAR
		IN :	BOOL;
		MANUAL :	BOOL;
		RST :	BOOL := FALSE;
		MIN_ONTIME :	TIME := T#10s;
		MIN_OFFTIME :	TIME := T#10s;
		RUN_EVERY :	TIME := T#10000m;
		PUMP :	BOOL;
		RUNTIME :	UDINT;
		CYCLES :	UDINT;
		func_block : ACTUATOR_PUMP_Block;
	END_VAR
	func_block.IN := IN;
	func_block.MANUAL := MANUAL;
	func_block.RST := RST ;
	func_block.MIN_ONTIME := MIN_ONTIME;
	func_block.MIN_OFFTIME := MIN_OFFTIME;
	func_block.RUN_EVERY := RUN_EVERY ;
	func_block();
	PUMP  := func_block.PUMP;
	RUNTIME  := func_block.RUNTIME;
	CYCLES  := func_block.CYCLES;
END_PROGRAM

CONFIGURATION Config0
	VAR_GLOBAL
		PLC_TICKS_PER_SEC :	INT;
		PLC_SYS_TICK_CNT :	DINT;
	END_VAR
  	RESOURCE Res0 ON PLC
    	TASK task0(INTERVAL := T#20ms,PRIORITY := 0);
    	PROGRAM instance0 WITH task0 : program0;
  	END_RESOURCE
END_CONFIGURATION

(* ---- ACTUATOR_UD.ST ---- *)
FUNCTION_BLOCK T_PLC_MS_block
	VAR_OUTPUT
		T_PLC_MS :	UDINT;
	END_VAR

	VAR_EXTERNAL
		PLC_TICKS_PER_SEC :	INT;
		PLC_SYS_TICK_CNT :	DINT;
	END_VAR

	VAR
		debug :	BOOL;(*Debug-Mode ON / OFF*)
		N :	INT;(*Debug-Faktor*)
		Offset :	UDINT;(*Debug-Offset*)
		temp :	DWORD := DWORD#1;(*Debug-Offset*)
		mode :	BOOL;(*modus*)
		faktor :	UDINT;(*Systemtakt-Faktor*)
		init :	BOOL;
		v_plc_ticks_per_sec :	UDINT;
		base :	UDINT := UDINT#1000;
	END_VAR

	IF init = FALSE THEN
		v_plc_ticks_per_sec := INT_TO_UDINT(PLC_TICKS_PER_SEC);
		IF v_plc_ticks_per_sec = UDINT#1024 THEN
			faktor := UDINT#1;
			mode := FALSE;
		ELSIF v_plc_ticks_per_sec > UDINT#0 THEN
			IF v_plc_ticks_per_sec <= base THEN
				faktor := base / v_plc_ticks_per_sec;
				mode := FALSE;
			ELSE
				faktor := v_plc_ticks_per_sec / base;
				mode := TRUE;
			END_IF;
		ELSE
			faktor := UDINT#1;
		END_IF;
		init := TRUE;
	END_IF;

	IF mode THEN
		T_PLC_MS := DINT_TO_UDINT(PLC_SYS_TICK_CNT) / faktor;
	ELSE
		T_PLC_MS := DINT_TO_UDINT(PLC_SYS_TICK_CNT) * faktor;
	END_IF;

	IF debug THEN
		T_PLC_MS := (DWORD_TO_UDINT(SHL(UDINT_TO_DWORD(T_PLC_MS),N) OR SHL(temp,N)) - UDINT#1) + Offset;
	END_IF;
END_FUNCTION_BLOCK

FUNCTION_BLOCK ACTUATOR_UD_Block

	VAR_INPUT
		UD :	BOOL;
		_ON :	BOOL;
		MANUAL :	BOOL;
		UP :	BOOL;
		DN :	BOOL;
		OFF :	BOOL;
		YUP_IN :	BOOL;
		YDN_IN :	BOOL;
		_TON :	TIME;
		TOFF :	TIME;
		OUT_RETURN :	BOOL;
	END_VAR

	VAR_OUTPUT
		YUP :	BOOL;
		YDN :	BOOL;
		STATUS :	BYTE;
	END_VAR

	VAR
		tx :	TIME;
		last :	TIME;
		init :	BOOL;
		T_PLC_MS :	T_PLC_MS_Block;
	END_VAR

	T_PLC_MS();
	tx:= UDINT_TO_TIME(T_PLC_MS.T_PLC_MS);

	IF NOT init THEN
		last := tx;
		init := TRUE;
	ELSIF off THEN
		Yup := FALSE;
		Ydn := FALSE;
		last := tx;
		status := BYTE#101;

	ELSIF ((Yup OR Ydn) AND tx - last < _TON) THEN RETURN;
	ELSIF NOT yup AND NOT ydn AND tx - last < toff THEN	RETURN;

	ELSIF manual THEN
		status := BYTE#102;
		IF yup AND NOT up OR ydn AND NOT dn THEN
			ydn := FALSE;
			yup := FALSE;
			last := tx;
		ELSIF UP AND NOT DN AND NOT OFF THEN
			Ydn := FALSE;
			Yup := TRUE;
			last := tx;
			status := BYTE#103;
		ELSIF DN AND NOT UP AND NOT OFF THEN
			Yup := FALSE;
			Ydn := TRUE;
			last := tx;
			status := BYTE#104;
		ELSE
			IF YUP OR YDN THEN LAST := tx; END_IF;
			Yup := FALSE;
			Ydn := FALSE;
		END_IF;

	ELSE
		IF yup AND NOT ud OR ydn AND UD THEN
			yup := FALSE;
			ydn := FALSE;
			last := tx;
		ELSIF Ud AND _ON AND NOT OFF THEN
			Ydn := FALSE;
			Yup := TRUE;
			last := tx;
			status := BYTE#111;

		ELSIF NOT UD AND _ON AND NOT OFF THEN
			Yup := FALSE;
			Ydn := TRUE;
			last := tx;
			status := BYTE#112;
		ELSE
			IF Yup OR Ydn THEN last := tx; END_IF;
			Yup := FALSE;
			Ydn := FALSE;
			status := BYTE#110;
		END_IF;
	END_IF;

	IF Ydn AND Yup_in AND out_return THEN
		Ydn := FALSE;
		status := BYTE#1;
	END_IF;
	IF Yup AND Ydn_in AND out_return THEN
		Yup := FALSE;
		status := BYTE#2;
	END_IF;

END_FUNCTION_BLOCK

PROGRAM program0
	VAR
		UD :	BOOL;
		_ON :	BOOL;
		MANUAL :	BOOL;
		UP :	BOOL;
		DN :	BOOL;
		OFF :	BOOL;
		YUP_IN :	BOOL;
		YDN_IN :	BOOL;
		_TON :	TIME;
		TOFF :	TIME;
		OUT_RETURN :	BOOL;
		YUP :	BOOL;
		YDN :	BOOL;
		STATUS :	BYTE;
		func_block : ACTUATOR_UD_Block;
	END_VAR
	func_block.UD := UD;
	func_block._ON := _ON;
	func_block.MANUAL := MANUAL ;
	func_block.UP := UP;
	func_block.DN := DN;
	func_block.OFF := OFF ;
	func_block.YUP_IN := YUP_IN;
	func_block.YDN_IN := YDN_IN;
	func_block._TON := _TON ;
	func_block.TOFF := TOFF;
	func_block.OUT_RETURN := OUT_RETURN;
	func_block();
	YUP  := func_block.YUP;
	YDN  := func_block.YDN;
	STATUS  := func_block.STATUS;
END_PROGRAM

CONFIGURATION Config0
	VAR_GLOBAL
		PLC_TICKS_PER_SEC :	INT;
		PLC_SYS_TICK_CNT :	DINT;
	END_VAR
  	RESOURCE Res0 ON PLC
    	TASK task0(INTERVAL := T#20ms,PRIORITY := 0);
    	PROGRAM instance0 WITH task0 : program0;
  	END_RESOURCE
END_CONFIGURATION

(* ---- AIN1.ST ---- *)
FUNCTION_BLOCK AIN1

	VAR_INPUT
		IN :	DWORD;
		SIGN_BIT :	INT := 255;
		ERROR_BIT :	INT := 255;
		ERROR_CODE_EN :	BOOL := FALSE;
		ERROR_CODE :	DWORD;
		OVERFLOW_BIT :	INT := 255;
		OVERFLOW_CODE_EN :	BOOL;
		OVERFLOW_CODE :	DWORD;
		BIT_0 :	INT;
		BIT_N :	INT := 31;
		OUT_MIN :	REAL;
		OUT_MAX :	REAL := 10.0;
		CODE_MIN :	DWORD;
		CODE_MAX :	DWORD := DWORD#16#FFFFFFFF;
		ERROR_OUTPUT :	REAL;
		OVERFLOW_OUTPUT :	REAL := 10.0;
	END_VAR

	VAR_OUTPUT
		OUT :	REAL;
		SIGN :	BOOL;
		ERROR :	BOOL;
		OVERFLOW :	BOOL;
	END_VAR

	VAR
		tB :	DWORD;
	END_VAR

	error := ((SHR(in,error_bit) AND DWORD#16#0000_0001) = DWORD#1) OR (error_code_en AND error_code = in);
	IF error THEN
		out := error_output;
		RETURN;
	END_IF;

	tb := SHR(SHL(in, 31 - bit_N), 31 - bit_N + Bit_0);

	overflow := ((SHR(in,overflow_bit) AND DWORD#16#0000_0001) = DWORD#1) OR (overflow_code_en AND overflow_code = in) OR (tb < code_min OR tb > code_max);
	IF overflow THEN
		out := overflow_output;
		RETURN;
	END_IF;

	sign := (SHR(in,sign_bit) AND DWORD#16#0000_0001) = DWORD#1;

	out := (UDINT_TO_REAL(DWORD_TO_UDINT(tb) - DWORD_TO_UDINT(code_min)) * (out_max - out_min) / UDINT_TO_REAL(DWORD_TO_UDINT(code_max) - DWORD_TO_UDINT(code_min)) + out_min);
	IF sign THEN out := out * -1.0; END_IF;

	(* extract error bit *)
	error := ((SHR(in,error_bit) AND DWORD#16#0000_0001) = DWORD#1) OR (error_code_en AND error_code = in);
	IF error THEN
		out := error_output;
		RETURN;
	END_IF;

	(* strip off the data input *)
	tb := SHR(SHL(in, 31 - bit_N), 31 - bit_N + Bit_0);

	(* extract overflow bit *)
	overflow := ((SHR(in,overflow_bit) AND DWORD#16#0000_0001) = DWORD#1) OR (overflow_code_en AND overflow_code = in) OR (tb < code_min OR tb > code_max);
	IF overflow THEN
		out := overflow_output;
		RETURN;
	END_IF;

	(* extract sign bit *)
	sign := (SHR(in,sign_bit) AND DWORD#16#0000_0001) = DWORD#1;

	(* convert in to out *)
	out := (UDINT_TO_REAL(DWORD_TO_UDINT(tb) - DWORD_TO_UDINT(code_min)) * (out_max - out_min) / UDINT_TO_REAL(DWORD_TO_UDINT(code_max) - DWORD_TO_UDINT(code_min)) + out_min);
	IF sign THEN out := out * - 1.0; END_IF;

END_FUNCTION_BLOCK

PROGRAM program0
  VAR
	IN               :	DWORD;
	SIGN_BIT         :	INT ;
	ERROR_BIT        :	INT ;
	ERROR_CODE_EN    :	BOOL ;
	ERROR_CODE       :	DWORD;
	OVERFLOW_BIT     :	INT ;
	OVERFLOW_CODE_EN :	BOOL;
	OVERFLOW_CODE    :	DWORD;
	BIT_0            :	INT;
	BIT_N            :	INT;
	OUT_MIN          :	REAL;
	OUT_MAX          :	REAL ;
	CODE_MIN         :	DWORD;
	CODE_MAX         :	DWORD ;
	ERROR_OUTPUT     :	REAL;
	OVERFLOW_OUTPUT  :	REAL ;

	OUT      :	REAL;
	SIGN     :	BOOL;
	ERROR    :	BOOL;
	OVERFLOW :	BOOL;

	func_block : AIN1;
  END_VAR
	func_block.IN               :=IN              ;
	func_block.SIGN_BIT         :=SIGN_BIT        ;
	func_block.ERROR_BIT        :=ERROR_BIT       ;
	func_block.ERROR_CODE_EN    :=ERROR_CODE_EN   ;
	func_block.ERROR_CODE       :=ERROR_CODE      ;
	func_block.OVERFLOW_BIT     :=OVERFLOW_BIT    ;
	func_block.OVERFLOW_CODE_EN :=OVERFLOW_CODE_EN;
	func_block.OVERFLOW_CODE    :=OVERFLOW_CODE   ;
	func_block.BIT_0            :=BIT_0           ;
	func_block.BIT_N            :=BIT_N           ;
	func_block.OUT_MIN          :=OUT_MIN         ;
	func_block.OUT_MAX          :=OUT_MAX         ;
	func_block.CODE_MIN         :=CODE_MIN        ;
	func_block.CODE_MAX         :=CODE_MAX        ;
	func_block.ERROR_OUTPUT     :=ERROR_OUTPUT    ;
	func_block.OVERFLOW_OUTPUT  :=OVERFLOW_OUTPUT ;

	func_block();
	OUT     := func_block.OUT     ;
	SIGN    := func_block.SIGN    ;
	ERROR   := func_block.ERROR   ;
	OVERFLOW:= func_block.OVERFLOW;
END_PROGRAM

CONFIGURATION Config0
  RESOURCE Res0 ON PLC
    TASK task0(INTERVAL := T#20ms,PRIORITY := 0);
    PROGRAM instance0 WITH task0 : program0;
  END_RESOURCE
END_CONFIGURATION
